(* IEC 61131-3 sources: JingjiangArm/moonboxpro_arm_8.4/Application/Application/任务列表/Main_Task, 12 files *)

(* ---- StErrParam_Use.st ---- *)
(*@CES
Name=StErrParam_Use
Type=Gvl
TypeGuid=2db5746d-d284-4425-9f7f-2663a34b0ebc
Guid=58394340-2af0-469d-907b-43e2b620f20c
HasDeclaration=True
HasImplementation=False
*)
{DECLARATION}
{attribute 'pack_mode' := '1'}
TYPE StErrParam_Use :(*这个是最终计算调整量需要的所有误差相关内容*)
STRUCT
	iErr_V: INT;(*纵向误差*)
	iErr_H: INT;(*横向误差*)
	iErr_V_Unprocessed	: INT;(*纵向误差-原始误差*)
	iErr_H_Unprocessed	: INT;(*横向误差-原始误差*)
	byIDX_V: BYTE;(*纵向索引*)
	byIDX_H: BYTE;(*横向索引*)
	byErrSts: BYTE;(*误差状态*)
	uiFSampleCounter:UINT;(*精采样数据计数*)
	iVerror_FollowPreUnit:INT;(*纵向跟踪前一色误差*)
	iVerror_Follow1Unit:INT;(*纵向跟踪第一色误差*)
	iHerror_FollowPreUnit :INT 	; (*横向跟前一色误差*)
	iHerror_Follow1Unit :INT 	;(*横向跟1色误差*)
	(*2025.9.16.094302*)
	iResult_VFollowpre_1stDerivate	: INT;(*YZJ计算误差*)
	//2025.11.13.105908||上传基线和峰值
	uiPeakValue_t1				: UINT;
	uiPeakValue_t2				: UINT;
	uiBaseUse_t1				: UINT;
	uiBaseUse_t2				: UINT;
	//2026.4.11.153149+2026.5.9.110438
	iErr_V_Display	: INT;(*纵向误差-显示平均处理*)
	iErr_H_Display	: INT;(*横向误差-原始误差*)

//2026.5.12.202228
	(*2026.5.10.150407/han.dp*)
	uiV_cam_raw: UINT;(*相机纵向原始误差*)
	iV_cam_pure: INT;(*相机纵向纯误差*)
	uiH_cam_raw: UINT;(*相机横向原始误差*)
	iH_cam_pure: INT;(*相机横向纯误差*)

END_STRUCT
END_TYPE

{IMPLEMENTATION}

(* ---- StTaskCycleDetection.st ---- *)
(*@CES
Name=StTaskCycleDetection
Type=Gvl
TypeGuid=2db5746d-d284-4425-9f7f-2663a34b0ebc
Guid=d17a89bb-f73c-4312-a6cf-f8b703e65793
HasDeclaration=True
HasImplementation=False
*)
{DECLARATION}
TYPE StTaskCycleDetection :
STRUCT
	xRstDetection			: BOOL;(* 复位测量 *)
	udiCycleCnt				: UDINT;(* 周期计数 *)
	xCalcIntervalEnabled	: BOOL;(* 计算间隔有效 *)
	tmTskIn					: TIME;(* 进入任务的时间戳 *)
	tmTskOut				: TIME;(* 离开任务的时间戳 *)
	tmTskIn_Prev			: TIME;(* 上次进入任务的时间戳 *)
	tmElapsed				: TIME;(* 任务消耗时间 *)
	tmElapsedMax			: TIME;(* 任务消耗时间最大 *)
	tmInterval				: TIME;(* 任务间隔 *)
	tmIntervalMax			: TIME;(* 任务间隔最大 *)
END_STRUCT
END_TYPE

{IMPLEMENTATION}

(* ---- KS_FlyMedian.st ---- *)
(*@CES
Name=KS_FlyMedian
Type=FunctionBlock
TypeGuid=6f9dac99-8de1-4efc-8465-68ac443b7d08
Guid=38054e60-5949-4eec-bd09-7b0f80079a4b
HasDeclaration=True
HasImplementation=True
*)
{DECLARATION}
FUNCTION KS_FlyMedian : REAL
(*中位数:与Python statistics.median语义一致——奇数取正中,偶数取中间两值的平均*)
(*插入排序会打乱入参缓冲区,窗口<=64,代价可忽略|Yang.zj+用于新飞点检测 2026.10.24.191149*)
VAR_INPUT
	pBuf	: POINTER TO REAL;(*缓冲区指针*)
	iCnt	: INT;			(*元素个数*)
END_VAR
VAR
	i		: INT;
	j		: INT;
	rTmp	: REAL;
END_VAR

{IMPLEMENTATION}
IF iCnt <= 0 THEN
	KS_FlyMedian:= 0.0;
	RETURN;
END_IF
FOR i:= 1 TO iCnt-1 DO(*插入排序*)
	rTmp:= pBuf[i];
	j:= i-1;
	WHILE (j >= 0) DO
		IF pBuf[j] > rTmp THEN
			pBuf[j+1]:= pBuf[j];
			j:= j-1;
		ELSE
			EXIT;
		END_IF
	END_WHILE
	pBuf[j+1]:= rTmp;
END_FOR
IF (iCnt MOD 2) = 1 THEN
	KS_FlyMedian:= pBuf[iCnt/2];
ELSE
	KS_FlyMedian:= (pBuf[iCnt/2-1] + pBuf[iCnt/2]) * 0.5;
END_IF

(* ---- KS_TskCycle_Begin.st ---- *)
(*@CES
Name=KS_TskCycle_Begin
Type=FunctionBlock
TypeGuid=6f9dac99-8de1-4efc-8465-68ac443b7d08
Guid=4df1a699-322b-4ad9-8d1d-9083be64c28d
HasDeclaration=True
HasImplementation=True
*)
{DECLARATION}
FUNCTION KS_TskCycle_Begin : INT
VAR_INPUT
	i_pstStTaskCycleDetection: POINTER TO StTaskCycleDetection;
END_VAR
VAR
	iResult: INT;
END_VAR
{IMPLEMENTATION}
iResult:= 0;
IF i_pstStTaskCycleDetection<>0 THEN
	i_pstStTaskCycleDetection^.tmTskIn:= TIME(); (* 进入的时间 *)
	i_pstStTaskCycleDetection^.udiCycleCnt:= i_pstStTaskCycleDetection^.udiCycleCnt+1; (* 进入一次就累计1次 *)
ELSE
	iResult:= -1;
END_IF
KS_TskCycle_Begin:= iResult;

(* ---- KS_TskCycle_End.st ---- *)
(*@CES
Name=KS_TskCycle_End
Type=FunctionBlock
TypeGuid=6f9dac99-8de1-4efc-8465-68ac443b7d08
Guid=379e6dd0-0b0c-44de-a9dc-120ed630a8f7
HasDeclaration=True
HasImplementation=True
*)
{DECLARATION}
FUNCTION KS_TskCycle_End : INT
VAR_INPUT
	i_pstStTaskCycleDetection: POINTER TO StTaskCycleDetection;
END_VAR
VAR
	iResult: INT;
END_VAR
{IMPLEMENTATION}
iResult:= 0;
IF i_pstStTaskCycleDetection<>0 THEN
	i_pstStTaskCycleDetection^.tmTskOut:= TIME(); (* 结束的时间 *)
	i_pstStTaskCycleDetection^.tmElapsed:= i_pstStTaskCycleDetection^.tmTskOut-i_pstStTaskCycleDetection^.tmTskIn; (* 算出本次耗时 *)
	IF i_pstStTaskCycleDetection^.tmElapsed>i_pstStTaskCycleDetection^.tmElapsedMax THEN (* 如果最高纪录有变化 *)
		i_pstStTaskCycleDetection^.tmElapsedMax:= i_pstStTaskCycleDetection^.tmElapsed;
	END_IF
	IF NOT i_pstStTaskCycleDetection^.xCalcIntervalEnabled THEN
		i_pstStTaskCycleDetection^.xCalcIntervalEnabled:= TRUE;
	ELSE
		i_pstStTaskCycleDetection^.tmInterval:= i_pstStTaskCycleDetection^.tmTskIn-i_pstStTaskCycleDetection^.tmTskIn_Prev; (* 周期间隔 *)
		IF i_pstStTaskCycleDetection^.tmInterval>i_pstStTaskCycleDetection^.tmIntervalMax THEN (* 如果周期间隔纪录有变化 *)
			i_pstStTaskCycleDetection^.tmIntervalMax:= i_pstStTaskCycleDetection^.tmInterval;
		END_IF
	END_IF

	i_pstStTaskCycleDetection^.tmTskIn_Prev:= i_pstStTaskCycleDetection^.tmTskIn; (* 上次进入的时间 *)

	IF i_pstStTaskCycleDetection^.xRstDetection THEN (* 重新计算周期的操作 *)
		i_pstStTaskCycleDetection^.xRstDetection:= FALSE;
		i_pstStTaskCycleDetection^.xCalcIntervalEnabled:= FALSE;
		i_pstStTaskCycleDetection^.tmElapsedMax:= T#0ms;
		i_pstStTaskCycleDetection^.tmIntervalMax:= T#0ms;
	END_IF
ELSE
	iResult:= -1;
END_IF

KS_TskCycle_End:= iResult;

(* ---- KS_UnPack_VisionERR.st ---- *)
(*@CES
Name=KS_UnPack_VisionERR
Type=FunctionBlock
TypeGuid=6f9dac99-8de1-4efc-8465-68ac443b7d08
Guid=46688986-88ab-493d-84a0-0feefd58abe3
HasDeclaration=True
HasImplementation=True
*)
{DECLARATION}
FUNCTION KS_UnPack_VisionERR : INT
VAR_INPUT
	i_wERR: WORD;(*接收到的误差值-加密数据*)
	i_pxFlag_valid: POINTER TO BOOL;(*bit15/有效标志*)
	i_pxFlag_update: POINTER TO BOOL;(*bit14/更新标志*)
	i_pxFlag_bitchk: POINTER TO BOOL;(*bit13/校验位*)
	i_piErr: POINTER TO INT;(*bit12~0/误差*)
END_VAR
VAR
	iRtn: INT := 0;(*默认0*)
END_VAR

{IMPLEMENTATION}
IF i_pxFlag_valid<>0 AND
	i_pxFlag_update<>0 AND
	i_pxFlag_bitchk<>0 AND
	i_piErr<>0 THEN
	iRtn:= 0;
	i_pxFlag_valid^:= WORD_TO_BOOL(SHR(i_wERR, 15) AND 16#1);
	i_pxFlag_update^:= WORD_TO_BOOL(SHR(i_wERR, 14) AND 16#1);
	i_pxFlag_bitchk^:= WORD_TO_BOOL(SHR(i_wERR, 13) AND 16#1);
	i_piErr^:= SHR(WORD_TO_INT(SHL(i_wERR, 3)), 3);
ELSE
	iRtn:= -1;
END_IF
KS_UnPack_VisionERR:= iRtn;

(* ---- KS_FB_AverageErr_Arc.st ---- *)
(*@CES
Name=KS_FB_AverageErr_Arc
Type=FunctionBlock
TypeGuid=6f9dac99-8de1-4efc-8465-68ac443b7d08
Guid=91f3b4d4-1a1f-49cc-9d09-db86b76ec74e
HasDeclaration=True
HasImplementation=True
*)
{DECLARATION}
FUNCTION_BLOCK KS_FB_AverageErr_Arc
VAR_INPUT
	i_xEn: BOOL;
	i_iErr: INT;(*输入的有效误差*)
	i_xErrValid: BOOL;(*误差有效性*)
	i_byAverageNum: BYTE;(*误差平均次数*)
END_VAR
VAR_OUTPUT
	o_xEn: BOOL;
	o_iErNo: INT;
	o_iErrResult: INT;
END_VAR
VAR
	rErrResult: REAL;(*误差平均使用的*)
	iBufferedIndexRd				: INT							;(*buffered array read index|*)
	iBufferedIndexWr				: INT							;(*buffered array write index|*)
	iPushedErrItemsAtLeast			: INT							;
	arErrorBuffered			: ARRAY [1..20] OF REAL						;
	iCountForSignalLost				: INT	;
	rSumTotal						: REAL;
	iIndex							: INT;
END_VAR

{IMPLEMENTATION}
o_xEn:= i_xEn;
o_iErNo:= 0;
IF i_xEn THEN
	IF i_byAverageNum>0 THEN
		rErrResult:= INT_TO_REAL(i_iErr);
		IF i_xErrValid THEN
			iBufferedIndexWr:= iBufferedIndexWr+1;
			IF iBufferedIndexWr>20 THEN
				iBufferedIndexWr:= iBufferedIndexWr-20;
			END_IF
			arErrorBuffered[iBufferedIndexWr]:= rErrResult;
			IF iPushedErrItemsAtLeast<i_byAverageNum THEN
				iPushedErrItemsAtLeast:= iPushedErrItemsAtLeast+1;
			ELSE
				IF i_byAverageNum>1 THEN
					iBufferedIndexRd:= iBufferedIndexWr;
					rSumTotal:= 0;
					FOR iIndex:=1 TO i_byAverageNum BY 1 DO
						rSumTotal:= rSumTotal+arErrorBuffered[iBufferedIndexRd];
						iBufferedIndexRd:= iBufferedIndexRd-1;
						IF iBufferedIndexRd<1 THEN
							iBufferedIndexRd:= iBufferedIndexRd+20;
						END_IF
					END_FOR
					rErrResult:= rSumTotal/i_byAverageNum;
				END_IF
			END_IF
			iCountForSignalLost:= 0;
			o_iErrResult:= REAL_TO_INT(rErrResult) ;
		ELSE(*连续丢失3幅就重新开始计算平均*)
			iCountForSignalLost:= 	iCountForSignalLost+1;
			IF 	iCountForSignalLost>3 THEN
				iBufferedIndexWr:= 0;
				iPushedErrItemsAtLeast:= 0;
			END_IF
			o_iErNo:= -1;
		END_IF
	ELSE
		o_iErrResult:= i_iErr;
	END_IF
END_IF

(* ---- KS_FB_GetError_Arc.st ---- *)
(*@CES
Name=KS_FB_GetError_Arc
Type=FunctionBlock
TypeGuid=6f9dac99-8de1-4efc-8465-68ac443b7d08
Guid=34f07fc4-d98c-4616-a827-05a7c8017d66
HasDeclaration=True
HasImplementation=True
*)
{DECLARATION}
FUNCTION_BLOCK KS_FB_GetError_Arc
VAR_INPUT
	i_xEn: BOOL;
	i_iUnitMax: INT;
	i_byGetErrMode: BYTE;(*获取误差方式，
	1：读取金刚来的误差
	2：读取月光宝盒/月光宝盒PRO来的误差
	*)
	i_aiAlarm_V: ARRAY [1..MAX_UNIT_NUM] OF INT;(*后续换成全局输入的变量*)
	i_aiAlarm_H: ARRAY [1..MAX_UNIT_NUM] OF INT;(*后续换成全局输入的变量*)
	i_aiAdjust_V: ARRAY [1..MAX_UNIT_NUM] OF INT;(*修正量*)
	i_aiAdjust_H: ARRAY [1..MAX_UNIT_NUM] OF INT;(*修正量*)

	i_abyAverageNum_V: ARRAY [1..MAX_UNIT_NUM] OF BYTE;(*误差平均次数*)
	i_abyAverageNum_H: ARRAY [1..MAX_UNIT_NUM] OF BYTE;(*误差平均次数*)
	//2026.4.11.150236 误差显示平均
	i_abyAverageNum_V_Display: ARRAY [1..MAX_UNIT_NUM] OF BYTE;(*误差显示平均次数*)
	i_abyAverageNum_H_Display: ARRAY [1..MAX_UNIT_NUM] OF BYTE;(*误差显示平均次数*)
	i_pstStSysParam								: POINTER TO StSysParam;
END_VAR
VAR_OUTPUT
	o_xEn: BOOL;
	o_iNoEr: INT;
	o_astStErrParam_Use: ARRAY [1..MAX_UNIT_NUM] OF StErrParam_Use;
END_VAR
VAR
	iN: INT;
	aiError_and_Sts_V: ARRAY [1..MAX_UNIT_NUM] OF INT;(*读取的来自金刚/月光宝盒PRO的误差及状态*)
	aiError_and_Sts_H: ARRAY [1..MAX_UNIT_NUM] OF INT;(*读取的来自金刚/月光宝盒PRO的误差及状态*)
	iTemp: WORD;
	aiError_V: ARRAY [1..MAX_UNIT_NUM] OF INT;(*处理完成后的纵向误差列表*)
	aiError_H: ARRAY [1..MAX_UNIT_NUM] OF INT;(*处理完成后的横向误差列表*)
	abyErrSts: ARRAY [1..MAX_UNIT_NUM] OF BYTE;(*处理完成后的纵横向误差状态*)
	abyIndex_V: ARRAY [1..MAX_UNIT_NUM] OF BYTE;(*处理完成后的索引*)
	abyIndex_H: ARRAY [1..MAX_UNIT_NUM] OF BYTE;(*处理完成后的索引*)
	axValid_V: ARRAY [1..MAX_UNIT_NUM] OF BOOL;(*误差有效性*)
	axValid_H: ARRAY [1..MAX_UNIT_NUM] OF BOOL;(*误差有效性*)
	axFlag_Refresh_V: ARRAY [1..MAX_UNIT_NUM] OF BOOL;(*误差刷新标志*)
	axFlag_Refresh_H: ARRAY [1..MAX_UNIT_NUM] OF BOOL;(*误差刷新标志*)
	axFlag_Check_V: ARRAY [1..MAX_UNIT_NUM] OF BOOL;(*误差校验位*)
	axFlag_Check_H: ARRAY [1..MAX_UNIT_NUM] OF BOOL;(*误差校验位*)
	axFlag_PreRefresh_V: ARRAY [1..MAX_UNIT_NUM] OF BOOL;(*误差有效性*)
	axFlag_PreRefresh_H: ARRAY [1..MAX_UNIT_NUM] OF BOOL;(*误差有效性*)
	afbKS_FB_PickOutFakePoint_V: ARRAY [1..MAX_UNIT_NUM] OF KS_FB_PickOutFakePoint;(*误差飞点处理*)
	afbKS_FB_PickOutFakePoint_H: ARRAY [1..MAX_UNIT_NUM] OF KS_FB_PickOutFakePoint;
	afbKS_FB_AverageErr_Arc_V: ARRAY [1..MAX_UNIT_NUM] OF KS_FB_AverageErr_Arc;(*误差平均处理*)
	afbKS_FB_AverageErr_Arc_H: ARRAY [1..MAX_UNIT_NUM] OF KS_FB_AverageErr_Arc;
	//2026.4.11.150050+
	afbKS_FB_AverageErr_Arc_V_Display: ARRAY [1..MAX_UNIT_NUM] OF KS_FB_AverageErr_Arc;(*误差平均处理@界面显示*)
	afbKS_FB_AverageErr_Arc_H_Display: ARRAY [1..MAX_UNIT_NUM] OF KS_FB_AverageErr_Arc;

	aiError_V_Res_Display: ARRAY [1..MAX_UNIT_NUM] OF INT;(*处理完成后的纵向显示误差列表*)
	aiError_H_Res_Display: ARRAY [1..MAX_UNIT_NUM] OF INT;(*处理完成后的横向显示误差列表*)
	//2026.5.9.110955
	axFakePoint_V: ARRAY [1..MAX_UNIT_NUM] OF BOOL;
	axFakePoint_H: ARRAY [1..MAX_UNIT_NUM] OF BOOL;

	aiError_V_Res: ARRAY [1..MAX_UNIT_NUM] OF INT;(*处理完成后的纵向误差列表*)
	aiError_H_Res: ARRAY [1..MAX_UNIT_NUM] OF INT;(*处理完成后的横向误差列表*)
	abyIndex_V_Pre: ARRAY [1..MAX_UNIT_NUM] OF BYTE;(*处理完成后的索引*)
	abyIndex_H_Pre: ARRAY [1..MAX_UNIT_NUM] OF BYTE;(*处理完成后的索引*)
	iUnitNR: INT;
	iStationId: INT;
	dwOFST2: DWORD;
	iRtn: INT;
	stStProtocol_PDU_Up_Rd: StParam_PDU_Up;
	pstStCMD_F05_: POINTER TO StPdu_Up_05;
	pbyTemp: POINTER TO BYTE;
	wCHK_Up_Calc: WORD;
	dwCheckSumVal: DWORD;
	abyBuf_PduCmd_rcv: ARRAY [1..MAX_PDU_CMD_BYTES_UP] OF BYTE; (* 2021.12.4.163129/hdp/读取 *)
	xtest: BOOL;
	aiResult_VFollowpre_1stDerivate: ARRAY [1..MAX_UNIT_NUM] OF INT;

	//alTime: ARRAY [1..10] OF LTIME;
	abyBuf_PduCmd_rcv_All: ARRAY [1..1000] OF BYTE;

	//新飞点剔除:每色组纵横各一个独立实例(总开关gc_xUseNewFlyRemove在GCL)|Yang.zj+用于新飞点检测 2026.10.24.191149
	afbKS_FlyRemove_V: ARRAY [1..MAX_UNIT_NUM] OF KS_FlyRemove;
	afbKS_FlyRemove_H: ARRAY [1..MAX_UNIT_NUM] OF KS_FlyRemove;
	aiError_V_Fly: ARRAY [1..MAX_UNIT_NUM] OF INT;(*剔除后送平均的纵向误差*)
	aiError_H_Fly: ARRAY [1..MAX_UNIT_NUM] OF INT;(*剔除后送平均的横向误差*)
	xFlyNewFrame: BOOL;(*本周期该色组是否来了新帧*)
	xFlyReset: BOOL;(*该色组剔除器复位请求*)
	aiFlyMarkModePre: ARRAY [1..MAX_UNIT_NUM] OF INT;(*上次色标排列模式*)
	abyFlySignalPre: ARRAY [1..MAX_UNIT_NUM] OF BYTE;(*上次RGB信号通道*)
	axFlyHorEnPre: ARRAY [1..MAX_UNIT_NUM] OF BOOL;(*上次横向开关*)
END_VAR

{IMPLEMENTATION}
o_xEn:= i_xEn;
o_iNoEr:= 0;
IF i_xEn THEN
	IF i_iUnitMax>0 THEN
	CASE i_byGetErrMode OF
			1:
				FOR iN:=1 TO i_iUnitMax BY 1 DO
					iTemp:= aiError_and_Sts_V[iN];
					axValid_V[iN]:= INT_TO_BOOL(iTemp AND 16#04);(*bit2:有效位*)
					axFlag_Refresh_V[iN]:= INT_TO_BOOL(iTemp AND 16#02);(*bit1:刷新位*)
					axFlag_Check_V[iN]:= INT_TO_BOOL(iTemp AND 16#01);(*bit0:校验位*)
					IF axFlag_PreRefresh_V[iN]<>axFlag_Refresh_V[iN] THEN	 	(*误差已刷新*)
						IF axValid_V[iN] THEN
							aiError_V[iN]:= SHR(iTemp,3);(*误差*)
						ELSE
							aiError_V[iN]:= gc_iValueReferToLost;
							abyErrSts[iN].1:= TRUE;(*纵向丢失*)
						END_IF
						abyIndex_V[iN]:= abyIndex_V[iN]+1;
					END_IF
					axFlag_PreRefresh_V[iN]:= axFlag_Refresh_V[iN];
					(*纵向误差处理完成*)
					iTemp:= aiError_and_Sts_H[iN];
					axValid_H[iN]:= INT_TO_BOOL(iTemp AND 16#04);(*bit2:有效位*)
					axFlag_Refresh_H[iN]:= INT_TO_BOOL(iTemp AND 16#02);(*bit1:刷新位*)
					axFlag_Check_H[iN]:= INT_TO_BOOL(iTemp AND 16#01);(*bit0:校验位*)
					IF axFlag_PreRefresh_H[iN]<>axFlag_Refresh_H[iN] THEN	 	(*误差已刷新*)
						IF axValid_H[iN] THEN
							aiError_H[iN]:= SHR(iTemp,3);(*误差*)
						ELSE
							aiError_H[iN]:= gc_iValueReferToLost;
							abyErrSts[iN].5:= TRUE;(*横向丢失*)
						END_IF
						abyIndex_H[iN]:= abyIndex_H[iN]+1;
					END_IF
					axFlag_PreRefresh_H[iN]:= axFlag_Refresh_H[iN];
					(*横向误差处理完成*)
				END_FOR
			2:
				//alTime[4] := LTIME();
				dwOFST2:= 0;
				iRtn := GTN_RN_UserPCRdLocalFPGA(
							1,1,
							0,//0,
							ADR(abyBuf_PduCmd_rcv_All),
							DWORD_TO_WORD(dwOFST2),
							KS_GetNumOfDwordUsed(INT_TO_DWORD(i_iUnitMax)*MAX_PDU_CMD_BYTES_DN));
				FOR iN:=1 TO i_iUnitMax BY 1 DO
					iUnitNR:= iN;(*通讯轴号也需要根据后续系统配置处理*)
					iStationId:= g_stStSysParam.stStSysParam_UnSave.aiStationList_UnitController[iN];(*2024.1.3.200541/+ *)
					IF KS_IsValidStationNR(iStationId) THEN
					(*读取从站即时上报的数据|每次32Bytes|*)
//2025.11.20.172237
//						dwOFST2 := MAX_PDU_CMD_BYTES_DN*(iUnitNR-1);
// 						dwOFST2.14:= TRUE;(* 绝对地址访问 *)
(*						iRtn := GTN_RN_UserPCRdLocalFPGA(1,1,
									0,//INT_TO_BYTE(iStationId),
									ADR(stStProtocol_PDU_Up_Rd),
									DWORD_TO_WORD(dwOFST2),
									15);//16448
									*)
// 						iRtn := GTN_RN_UserPCRdLocalFPGA(
// 									ADR(stStProtocol_PDU_Up_Rd),
// 									0,//INT_TO_BYTE(iStationId),
// 									DWORD_TO_WORD(dwOFST2),
// 									15);//16448

//2025.11.20.172246
//						iRtn := GTN_RN_UserPCRdLocalFPGA(
// 									1,1,
// 									0,//0,
// 									ADR(abyBuf_PduCmd_rcv),
// 									DWORD_TO_WORD(dwOFST2),
// 									15);//16448
					dwOFST2 := MAX_PDU_CMD_BYTES_DN*(iUnitNR-1);

					SysMemCpy(ADR(stStProtocol_PDU_Up_Rd),ADR(abyBuf_PduCmd_rcv_All)+dwOFST2,SIZEOF(stStProtocol_PDU_Up_Rd));
					(*检查命令|*)
						pstStCMD_F05_:=0;

						pbyTemp:= ADR(stStProtocol_PDU_Up_Rd.byPkgId);
						wCHK_Up_Calc:= KS_CRC(pbyTemp, 46, ADR(dwCheckSumVal));(*51是wCHK之前的数据长度*)
						IF wCHK_Up_Calc=stStProtocol_PDU_Up_Rd.wCHK THEN (*CRC校验通过*)
							CASE stStProtocol_PDU_Up_Rd.byPkgId OF
								5:
								pstStCMD_F05_:= ADR(stStProtocol_PDU_Up_Rd.abyPayload);
								IF pstStCMD_F05_<>0 THEN
									aiError_V[iN]:= stStProtocol_PDU_Up_Rd.iErr_V_Raw;
									aiError_H[iN]:= stStProtocol_PDU_Up_Rd.iErr_H_Raw;
									abyIndex_V[iN]:= stStProtocol_PDU_Up_Rd.byIDX_V;
									abyIndex_H[iN]:= stStProtocol_PDU_Up_Rd.byIDX_H;
									IF aiError_V[iN]=gc_iValueReferToLost THEN
										abyErrSts[iN].1:= TRUE;(*纵向丢失*)
									ELSE
										axValid_V[iN]:= TRUE;
									END_IF
									IF aiError_H[iN]=gc_iValueReferToLost THEN
										abyErrSts[iN].5:= TRUE;(*横向丢失*)
									ELSE
										axValid_H[iN]:= TRUE;
									END_IF
									o_astStErrParam_Use[iN].iResult_VFollowpre_1stDerivate:=
											pstStCMD_F05_^.iResult_VFollowpre_1stDerivate;
									aiResult_VFollowpre_1stDerivate[iN]:=
											pstStCMD_F05_^.iResult_VFollowpre_1stDerivate;
									//2025.11.13.110235上传基线和峰值
									o_astStErrParam_Use[iN].uiBaseUse_t1:= pstStCMD_F05_^.uiBaseUse_t1;
									o_astStErrParam_Use[iN].uiBaseUse_t2:= pstStCMD_F05_^.uiBaseUse_t2;
									o_astStErrParam_Use[iN].uiPeakValue_t1:= pstStCMD_F05_^.uiPeakValue_t1;
									o_astStErrParam_Use[iN].uiPeakValue_t2:= pstStCMD_F05_^.uiPeakValue_t2;
								//2026.5.9.110642
									i_pstStSysParam^.astStRSV_UnitParam_UnSave[iN].iCurLabelPos:= pstStCMD_F05_^.iCurLabelPos;(*本色三角标位置，点数*)
									i_pstStSysParam^.astStRSV_UnitParam_UnSave[iN].iPreLabelPos:= pstStCMD_F05_^.iPreLabelPos;(*前色三角标位置，点数*)
									i_pstStSysParam^.astStRSV_UnitParam_UnSave[iN].byFlag_CommFromSlave:= pstStCMD_F05_^.byFlag_CommFromSlave;(*bit0 xFlag_FindFirstSuccess;bit1 xFlag_FindPreSuccess*)
									i_pstStSysParam^.astStRSV_UnitParam_UnSave[iN].xFlag_FindFirstSuccess:= i_pstStSysParam^.astStRSV_UnitParam_UnSave[iN].byFlag_CommFromSlave.0;
									i_pstStSysParam^.astStRSV_UnitParam_UnSave[iN].xFlag_FindPreSuccess:= i_pstStSysParam^.astStRSV_UnitParam_UnSave[iN].byFlag_CommFromSlave.1;
									i_pstStSysParam^.astStRSV_UnitParam_UnSave[iN].byDetectedSignalCount:= pstStCMD_F05_^.byDetectedSignalCount;(*当前检测到色标个数*)
									i_pstStSysParam^.astStRSV_UnitParam_UnSave[iN].byMarkStep:= pstStCMD_F05_^.byMarkStep;(*当前全自动套印步骤*)
									i_pstStSysParam^.astStRSV_UnitParam_UnSave[iN].rGateSignalWidth_R:= BYTE_TO_REAL (pstStCMD_F05_^.byWidthRS) /10.0;(*粗采样计算波形宽度*)

								END_IF
							END_CASE
						END_IF
					END_IF
				END_FOR

			ELSE
			(*其他状态时，就先按丢失处理*)
				FOR iN:=1 TO MAX_UNIT_NUM BY 1 DO
					aiError_V[iN]:= gc_iValueReferToLost;
					aiError_H[iN]:= gc_iValueReferToLost;
					abyErrSts[iN].1:= TRUE;(*纵向丢失*)
					abyErrSts[iN].5:= TRUE;(*横向丢失*)
				END_FOR
		END_CASE

		(*从这里开始进行误差处理-飞点和平均*)
		(*飞点处理*)

		(*FOR iN:=1 TO MAX_UNIT_NUM BY 1 DO
			IF abyIndex_V_Pre[iN]<>abyIndex_V[iN] AND abyIndex_H_Pre[iN]<>abyIndex_H[iN] THEN
				abyErrSts[iN]:= 0;
				axValid_V[iN]:= FALSE;
				axValid_H[iN]:= FALSE;
				IF aiError_V[iN]=gc_iValueReferToLost THEN
					abyErrSts[iN].1:= TRUE;(*纵向丢失*)
				ELSE
					axValid_V[iN]:= TRUE;
				END_IF
				IF aiError_H[iN]=gc_iValueReferToLost THEN
					abyErrSts[iN].5:= TRUE;(*横向丢失*)
				ELSE
					axValid_H[iN]:= TRUE;
				END_IF
				o_astStErrParam_Use[iN].iResult_VFollowpre_1stDerivate:=
						aiResult_VFollowpre_1stDerivate[iN];

				o_astStErrParam_Use[iN].byIDX_V:= abyIndex_V[iN];
				o_astStErrParam_Use[iN].byIDX_H:= abyIndex_H[iN];
	//2026.02.08.195855
				(*平均处理*)
				afbKS_FB_AverageErr_Arc_V[iN](
					i_xEn:= TRUE,
					i_iErr:= aiError_V[iN],
					i_xErrValid:= axValid_V[iN],(*2025.01.03.110017*)
					i_byAverageNum:= i_abyAverageNum_V[iN],
					o_iErrResult=>aiError_V_Res[iN]);
				axFakePoint_V[iN]:= FALSE;

				afbKS_FB_PickOutFakePoint_V[iN](
					i_xIsValidError:= axValid_V[iN],
					i_iError_0_01mm:= aiError_V_Res[iN],
					i_iVariationBaseValue:= 50,(*2025.01.03.110017*)
					i_iBoundaryError_0_01mm:= 20,
					i_iErrorLevel_0_01mm:= 25,
					i_iVariationVariationMin:= 5,
					i_iVariationVariationMax:= 50,
					o_xFakeIsConfirmed=> axFakePoint_V[iN]);
	//2026.02.08.195945
				afbKS_FB_AverageErr_Arc_H[iN](
					i_xEn:= TRUE,
					i_iErr:= aiError_H[iN],
					i_xErrValid:= axValid_H[iN],(*2025.01.03.110017*)
					i_byAverageNum:= i_abyAverageNum_H[iN],
					o_iErrResult=>aiError_H_Res[iN]);
				axFakePoint_H[iN]:= FALSE;

				afbKS_FB_PickOutFakePoint_H[iN](
					i_xIsValidError:= axValid_H[iN],
					i_iError_0_01mm:= aiError_H_Res[iN],
					i_iVariationBaseValue:= 50,
					i_iBoundaryError_0_01mm:= 20,
					i_iErrorLevel_0_01mm:= 25,
					i_iVariationVariationMin:= 5,
					i_iVariationVariationMax:= 50,
					o_xFakeIsConfirmed=> axFakePoint_H[iN]);

				//显示平均@2026.4.11.150119+
				afbKS_FB_AverageErr_Arc_V_Display[iN](
					i_xEn:= TRUE,
					i_iErr:= aiError_V[iN],
					i_xErrValid:= axValid_V[iN],(*2025.01.03.110017*)
					i_byAverageNum:= i_abyAverageNum_V_Display[iN],
					o_iErrResult=>aiError_V_Res_Display[iN]);

				afbKS_FB_AverageErr_Arc_H_Display[iN](
					i_xEn:= TRUE,
					i_iErr:= aiError_H[iN],
					i_xErrValid:= axValid_H[iN],(*2025.01.03.110017*)
					i_byAverageNum:= i_abyAverageNum_H_Display[iN],
					o_iErrResult=>aiError_H_Res_Display[iN]);

			END_IF*)
		FOR iN:=1 TO MAX_UNIT_NUM BY 1 DO
			(*新飞点剔除:误差平均之前对原始逐帧误差剔除,成熟账本时为外推 P 并刷锁存，否则锁存,必须先剔除再平均,否则飞点被N幅平均稀释后可能低于门限漏掉*)
			(*总开关gc_xUseNewFlyRemove在GCL,置FALSE并重编译即回退旧逻辑;飞点/暂缓帧置axFakePoint_V/H(byErrSts.2/6),阶跃(真实变化)不置位|Yang.zj+用于新飞点检测 2026.10.24.191149*)
			IF gc_xUseNewFlyRemove THEN
				xFlyNewFrame:= (abyIndex_V_Pre[iN]<>abyIndex_V[iN]) AND (abyIndex_H_Pre[iN]<>abyIndex_H[iN]);
				(*工况切换检测:色标排列模式/RGB信号通道/横向开关任一变化,该色组剔除器可信历史不可信,复位重新暖机*)
				xFlyReset:= FALSE;
				IF i_pstStSysParam<>0 THEN
					IF (aiFlyMarkModePre[iN]<>i_pstStSysParam^.astStUnitParam_Save[iN].iMarkArrangeMode)
						OR (abyFlySignalPre[iN]<>i_pstStSysParam^.astStUnitParam_Save[iN].bySignalSelect)
						OR (axFlyHorEnPre[iN]<>i_pstStSysParam^.astStUnitParam_Save[iN].dwFlag_Ctl.0) THEN
						aiFlyMarkModePre[iN]:= i_pstStSysParam^.astStUnitParam_Save[iN].iMarkArrangeMode;
						abyFlySignalPre[iN]:= i_pstStSysParam^.astStUnitParam_Save[iN].bySignalSelect;
						axFlyHorEnPre[iN]:= i_pstStSysParam^.astStUnitParam_Save[iN].dwFlag_Ctl.0;
						xFlyReset:= TRUE;
					END_IF
				END_IF
				afbKS_FlyRemove_V[iN](
					i_iErr:= aiError_V[iN],
					i_xErrValid:= xFlyNewFrame AND (aiError_V[iN]<>gc_iValueReferToLost),
					i_xLost:= xFlyNewFrame AND (aiError_V[iN]=gc_iValueReferToLost),
					i_xReset:= xFlyReset,
					o_iErrResult=> aiError_V_Fly[iN],
					o_xFake=> axFakePoint_V[iN]);
				afbKS_FlyRemove_H[iN](
					i_iErr:= aiError_H[iN],
					i_xErrValid:= xFlyNewFrame AND (aiError_H[iN]<>gc_iValueReferToLost),
					i_xLost:= xFlyNewFrame AND (aiError_H[iN]=gc_iValueReferToLost),
					i_xReset:= xFlyReset,
					o_iErrResult=> aiError_H_Fly[iN],
					o_xFake=> axFakePoint_H[iN]);
			ELSE
				aiError_V_Fly[iN]:= aiError_V[iN];(*旧路径:不剔除,原值送平均*)
				aiError_H_Fly[iN]:= aiError_H[iN];
			END_IF
			IF abyIndex_V_Pre[iN]<>abyIndex_V[iN] AND abyIndex_H_Pre[iN]<>abyIndex_H[iN] THEN
				abyErrSts[iN]:= 0;
				axValid_V[iN]:= FALSE;
				axValid_H[iN]:= FALSE;
				IF aiError_V[iN]=gc_iValueReferToLost THEN
					abyErrSts[iN].1:= TRUE;(*纵向丢失*)
				ELSE
					axValid_V[iN]:= TRUE;
				END_IF
				IF aiError_H[iN]=gc_iValueReferToLost THEN
					abyErrSts[iN].5:= TRUE;(*横向丢失*)
				ELSE
					axValid_H[iN]:= TRUE;
				END_IF
				o_astStErrParam_Use[iN].iResult_VFollowpre_1stDerivate:=
						aiResult_VFollowpre_1stDerivate[iN];

				o_astStErrParam_Use[iN].byIDX_V:= abyIndex_V[iN];
				o_astStErrParam_Use[iN].byIDX_H:= abyIndex_H[iN];
//2026.02.08.195855
				(*平均处理*)
				afbKS_FB_AverageErr_Arc_V[iN](
					i_xEn:= TRUE,
					i_iErr:= aiError_V_Fly[iN],(*新飞点:喂剔除后的值|Yang.zj+用于新飞点检测 2026.10.24.191149*)
					i_xErrValid:= axValid_V[iN],(*2025.01.03.110017*)
					i_byAverageNum:= i_abyAverageNum_V[iN],
					o_iErrResult=>aiError_V_Res[iN]);
				IF NOT gc_xUseNewFlyRemove THEN(*旧飞点判断:新算法启用时整块跳过|Yang.zj+用于新飞点检测 2026.10.24.191149*)
				axFakePoint_V[iN]:= FALSE;

				afbKS_FB_PickOutFakePoint_V[iN](
					i_xIsValidError:= axValid_V[iN],
					i_iError_0_01mm:= aiError_V_Res[iN],
					i_iVariationBaseValue:= 50,(*2025.01.03.110017*)
					i_iBoundaryError_0_01mm:= 20,
					i_iErrorLevel_0_01mm:= 25,
					i_iVariationVariationMin:= 5,
					i_iVariationVariationMax:= 50,
					o_xFakeIsConfirmed=> axFakePoint_V[iN]);
				END_IF
//2026.02.08.195945
				afbKS_FB_AverageErr_Arc_H[iN](
					i_xEn:= TRUE,
					i_iErr:= aiError_H_Fly[iN],(*新飞点:喂剔除后的值|Yang.zj+用于新飞点检测 2026.10.24.191149*)
					i_xErrValid:= axValid_H[iN],(*2025.01.03.110017*)
					i_byAverageNum:= i_abyAverageNum_H[iN],
					o_iErrResult=>aiError_H_Res[iN]);
				IF NOT gc_xUseNewFlyRemove THEN(*旧飞点判断:新算法启用时整块跳过|Yang.zj+用于新飞点检测 2026.10.24.191149*)
				axFakePoint_H[iN]:= FALSE;

				afbKS_FB_PickOutFakePoint_H[iN](
					i_xIsValidError:= axValid_H[iN],
					i_iError_0_01mm:= aiError_H_Res[iN],
					i_iVariationBaseValue:= 50,
					i_iBoundaryError_0_01mm:= 20,
					i_iErrorLevel_0_01mm:= 25,
					i_iVariationVariationMin:= 5,
					i_iVariationVariationMax:= 50,
					o_xFakeIsConfirmed=> axFakePoint_H[iN]);
				END_IF

				//显示平均@2026.4.11.150119+
				afbKS_FB_AverageErr_Arc_V_Display[iN](
					i_xEn:= TRUE,
					i_iErr:= aiError_V_Fly[iN],(*新飞点:喂剔除后的值|Yang.zj+用于新飞点检测 2026.10.24.191149*)
					i_xErrValid:= axValid_V[iN],(*2025.01.03.110017*)
					i_byAverageNum:= i_abyAverageNum_V_Display[iN],
					o_iErrResult=>aiError_V_Res_Display[iN]);

				afbKS_FB_AverageErr_Arc_H_Display[iN](
					i_xEn:= TRUE,
					i_iErr:= aiError_H_Fly[iN],(*新飞点:喂剔除后的值|Yang.zj+用于新飞点检测 2026.10.24.191149*)
					i_xErrValid:= axValid_H[iN],(*2025.01.03.110017*)
					i_byAverageNum:= i_abyAverageNum_H_Display[iN],
					o_iErrResult=>aiError_H_Res_Display[iN]);
			END_IF
			(*到这里误差的飞点和平均都处理完了，该处理其他东西了*)
			o_astStErrParam_Use[iN].iErr_V_Unprocessed:= aiError_V[iN];(*原始误差*)
			o_astStErrParam_Use[iN].iErr_H_Unprocessed:= aiError_H[iN];
			o_astStErrParam_Use[iN].byErrSts:= 0;
			o_astStErrParam_Use[iN].byErrSts:= abyErrSts[iN];(*现在的状态*)

//2026.5.9.110835处理一下显示平均相关
			IF NOT o_astStErrParam_Use[iN].byErrSts.1 THEN(*纵向未丢失*)
				o_astStErrParam_Use[iN].iErr_V:= aiError_V_Res[iN]-i_aiAdjust_V[iN];
				//2026.4.11.150603+
				o_astStErrParam_Use[iN].iErr_V_Display:= aiError_V_Res_Display[iN]-i_aiAdjust_V[iN];
				IF axFakePoint_V[iN] THEN(*飞点*)
					o_astStErrParam_Use[iN].byErrSts.2:= TRUE;
				END_IF
				(*报警标志检查*)
				//IF ABS(o_astStErrParam_Use[iN].iErr_V)>ABS(i_aiAlarm_V[iN]) THEN
				IF ABS(o_astStErrParam_Use[iN].iErr_V_Display)>ABS(i_aiAlarm_V[iN]) THEN
					o_astStErrParam_Use[iN].byErrSts.0:= TRUE;
				END_IF
			ELSE
				o_astStErrParam_Use[iN].iErr_V:= gc_iValueReferToLost;
				o_astStErrParam_Use[iN].iErr_V_Display:= gc_iValueReferToLost;
			END_IF
			IF NOT o_astStErrParam_Use[iN].byErrSts.5 THEN(*横向未丢失*)
				o_astStErrParam_Use[iN].iErr_H:= aiError_H_Res[iN]-i_aiAdjust_H[iN];(*处理完的误差-修正量*)
				//2026.4.11.150603+
				o_astStErrParam_Use[iN].iErr_H_Display:= aiError_H_Res_Display[iN]-i_aiAdjust_H[iN];
				IF axFakePoint_H[iN] THEN(*飞点*)
					o_astStErrParam_Use[iN].byErrSts.6:= TRUE;
				END_IF
				(*报警标志检查*)
				//IF ABS(o_astStErrParam_Use[iN].iErr_H)>ABS(i_aiAlarm_H[iN]) THEN
				IF ABS(o_astStErrParam_Use[iN].iErr_H_Display)>ABS(i_aiAlarm_H[iN]) THEN
					o_astStErrParam_Use[iN].byErrSts.4:= TRUE;
				END_IF
			ELSE
				o_astStErrParam_Use[iN].iErr_H:= gc_iValueReferToLost;
				//2026.4.11.150603+
				o_astStErrParam_Use[iN].iErr_H_Display:= gc_iValueReferToLost;
			END_IF
			abyIndex_V_Pre[iN]:= abyIndex_V[iN];
			abyIndex_H_Pre[iN]:= abyIndex_H[iN];
		END_FOR
	END_IF
END_IF

(* ---- KS_FB_GetError_Arc_1.st ---- *)
(*@CES
Name=KS_FB_GetError_Arc_1
Type=FunctionBlock
TypeGuid=6f9dac99-8de1-4efc-8465-68ac443b7d08
Guid=a8fc5d1b-180f-4776-912e-45955a246124
HasDeclaration=True
HasImplementation=True
*)
{DECLARATION}
FUNCTION_BLOCK KS_FB_GetError_Arc_1
VAR_INPUT
	i_xEn: BOOL;(*该功能的使能条件*)
	i_iUnitMax: INT;(*有效色组范围1..MAX_UNIT_NUM*)
	i_abyGetErrMode: ARRAY [1..MAX_UNIT_NUM] OF BYTE;
	(*2026.5.10.102830/han.dp/修正接口定义方式:
	bit0 月光宝盒PRO误差源,1有效
	bit1 金刚误差源,1有效
	bit4 相机安装方向-反向/2026.5.24.173347/han.dp
	bit5 逆序/2026.5.24.173354/han.dp
	bit7 用于标记有效位标志; =0表示bit0有效,以月光宝盒PRO的误差作为调整依据; =1表示bit1有效,以金刚误差作为调整参考;
	--------------------------------------------------
	举例:
	* 16#01来自月光宝盒PRO;
	* 16#82来自视觉,并作为调整依据;
	* 16#03金刚和月光宝盒PRO误差都读,但只以月光宝盒PRO的误差作为调整依据;
	* 16#83金刚和月光宝盒PRO误差都读,但只以金刚的误差作为调整依据;
	*)
	i_aiAlarm_V: ARRAY [1..MAX_UNIT_NUM] OF INT;(*后续换成全局输入的变量*)
	i_aiAlarm_H: ARRAY [1..MAX_UNIT_NUM] OF INT;(*后续换成全局输入的变量*)
	i_aiAdjust_V: ARRAY [1..MAX_UNIT_NUM] OF INT;(*修正量*)
	i_aiAdjust_H: ARRAY [1..MAX_UNIT_NUM] OF INT;(*修正量*)
	i_abyAverageNum_V: ARRAY [1..MAX_UNIT_NUM] OF BYTE;(*误差平均次数*)
	i_abyAverageNum_H: ARRAY [1..MAX_UNIT_NUM] OF BYTE;(*误差平均次数*)
	(*统一注释0916+2026.4.11.150236 误差显示平均*)
	i_abyAverageNum_V_Display: ARRAY [1..MAX_UNIT_NUM] OF BYTE;(*误差显示平均次数*)
	i_abyAverageNum_H_Display: ARRAY [1..MAX_UNIT_NUM] OF BYTE;(*误差显示平均次数*)
	i_pstStSysParam								: POINTER TO StSysParam;
	i_dwKSMatrixMark: DWORD;(*2026.5.24.173538/han.dp/科赛矩阵色标描述/高16bit和低16bit分别为ab值*)
END_VAR
VAR_OUTPUT
	o_xEno: BOOL;
	o_iErNo: INT;
	o_astStErrParam_Use: ARRAY [1..MAX_UNIT_NUM] OF StErrParam_Use;
	o_stSystimeElapsed: SYSTIME;(*2026.5.24.152004/han.dp*)
END_VAR
VAR
	xInitialized_Ref_KSMatrixMark: BOOL := FALSE;
	abyGetErrMode_Ref: ARRAY [1..MAX_UNIT_NUM] OF BYTE := [0];
	dwKSMatrixMark_Ref: DWORD := 0;
	aiRef_KSMatrixMark: ARRAY [1..MAX_UNIT_NUM,1..2] OF INT;(*16色色标的参考位置*)
	wKSMatrixMark_Hword: WORD;
	wKSMatrixMark_Lword: WORD;

	iN: INT;
	aiError_and_Sts_V: ARRAY [1..MAX_UNIT_NUM] OF INT;(*读取的来自金刚/月光宝盒PRO的误差及状态*)
	aiError_and_Sts_H: ARRAY [1..MAX_UNIT_NUM] OF INT;(*读取的来自金刚/月光宝盒PRO的误差及状态*)
	iTemp: WORD;

(*deprecated@2026.5.28.172423/han.dp
	axFlag_Refresh_V: ARRAY [1..MAX_UNIT_NUM] OF BOOL;(*误差刷新标志*)
	axFlag_Refresh_H: ARRAY [1..MAX_UNIT_NUM] OF BOOL;(*误差刷新标志*)
	axFlag_Check_V: ARRAY [1..MAX_UNIT_NUM] OF BOOL;(*误差校验位*)
	axFlag_Check_H: ARRAY [1..MAX_UNIT_NUM] OF BOOL;(*误差校验位*)
	axFlag_PreRefresh_V: ARRAY [1..MAX_UNIT_NUM] OF BOOL;(*误差有效性*)
	axFlag_PreRefresh_H: ARRAY [1..MAX_UNIT_NUM] OF BOOL;(*误差有效性*)
*)	afbKS_FB_PickOutFakePoint_V: ARRAY [1..MAX_UNIT_NUM] OF KS_FB_PickOutFakePoint;(*误差飞点处理*)
	afbKS_FB_PickOutFakePoint_H: ARRAY [1..MAX_UNIT_NUM] OF KS_FB_PickOutFakePoint;
	afbKS_FB_AverageErr_Arc_V: ARRAY [1..MAX_UNIT_NUM] OF KS_FB_AverageErr_Arc;(*误差平均处理*)
	afbKS_FB_AverageErr_Arc_H: ARRAY [1..MAX_UNIT_NUM] OF KS_FB_AverageErr_Arc;
	axFakePoint_V: ARRAY [1..MAX_UNIT_NUM] OF BOOL := [MAX_UNIT_NUM(FALSE)];
	axFakePoint_H: ARRAY [1..MAX_UNIT_NUM] OF BOOL := [MAX_UNIT_NUM(FALSE)];

	aiError_V_Res: ARRAY [1..MAX_UNIT_NUM] OF INT := [MAX_UNIT_NUM(0)];(*处理完成后的纵向误差列表*)
	aiError_H_Res: ARRAY [1..MAX_UNIT_NUM] OF INT := [MAX_UNIT_NUM(0)];(*处理完成后的横向误差列表*)
	abyIndex_V_Pre: ARRAY [1..MAX_UNIT_NUM] OF BYTE := [MAX_UNIT_NUM(0)];(*处理完成后的索引*)
	abyIndex_H_Pre: ARRAY [1..MAX_UNIT_NUM] OF BYTE := [MAX_UNIT_NUM(0)];(*处理完成后的索引*)

	iUnitNR: INT;
	iStationId: INT;
	dwOFST2: DWORD;

	iRtn: INT;
	stStProtocol_PDU_Up_Rd: StParam_PDU_Up;
	pstStCMD_F05_: POINTER TO StPdu_Up_05;
	pbyTemp: POINTER TO BYTE;
	wCHK_Up_Calc: WORD;
	dwCheckSumVal: DWORD;
(*	abyBuf_PduCmd_rcv: ARRAY [1..MAX_PDU_CMD_BYTES_UP] OF BYTE; (* 2021.12.4.163129/hdp/读取 *)*)
(*	xtest: BOOL;*)
	aiResult_VFollowpre_1stDerivate: ARRAY [1..MAX_UNIT_NUM] OF INT := [MAX_UNIT_NUM(0)];

	(*统一注释0916+alTime: ARRAY [1..10] OF LTIME;*)
	abyBuf_PduCmd_rcv_All: ARRAY [1..1000] OF BYTE;

	(*start___@2026.5.10.135832/han.dp
	视觉误差相关的补充变量*)
	adwErrMix_RdVision: ARRAY [1..MAX_UNIT_NUM] OF DWORD := [0];(*来自视觉的复合误差*)
	aiRtnMatrix: ARRAY [1..MAX_UNIT_NUM,1..2] OF INT := [0];(*处理误差解析的返回值矩阵*)
	aiErr_v_pure: ARRAY [1..MAX_UNIT_NUM] OF INT := [0];(*纵向实际误差/从金刚传来/未处理物理坐标系*)
	aiErr_h_pure: ARRAY [1..MAX_UNIT_NUM] OF INT := [0];(*横向实际误差/从金刚传来/未处理物理坐标系*)
(*	adwERR_VisionGave: ARRAY [1..MAX_UNIT_NUM] OF DWORD := [0];(*纵横向误差在一起*)*)

	axFlag_valid_v_tmp: ARRAY [1..MAX_UNIT_NUM] OF BOOL := [MAX_UNIT_NUM(FALSE)];(*纵向有效标志*)
	axFlag_update_v_tmp: ARRAY [1..MAX_UNIT_NUM] OF BOOL := [MAX_UNIT_NUM(FALSE)];(*纵向更新标志*)
	axFlag_update_v_rec: ARRAY [1..MAX_UNIT_NUM] OF BOOL := [MAX_UNIT_NUM(FALSE)];(*纵向上次更新标志*)
	axFlag_bitchk_v_tmp: ARRAY [1..MAX_UNIT_NUM] OF BOOL := [MAX_UNIT_NUM(FALSE)];(*纵向校验位*)

	axFlag_valid_h_tmp: ARRAY [1..MAX_UNIT_NUM] OF BOOL := [MAX_UNIT_NUM(FALSE)];(*横向有效标志*)
	axFlag_update_h_tmp: ARRAY [1..MAX_UNIT_NUM] OF BOOL := [MAX_UNIT_NUM(FALSE)];(*横向更新标志*)
	axFlag_update_h_rec: ARRAY [1..MAX_UNIT_NUM] OF BOOL := [MAX_UNIT_NUM(FALSE)];(*横向上次更新标志*)
	axFlag_bitchk_h_tmp: ARRAY [1..MAX_UNIT_NUM] OF BOOL := [MAX_UNIT_NUM(FALSE)];(*横向校验位*)

	pawErr_tmp: POINTER TO ARRAY [1..2] OF WORD := 0;
	(*___end@2026.5.10.135850*)

	stSystimeDelta,stSystimeStart,stSystimeEnd:SYSTIME;(*获取us时间差*)
	abyVisionErrIdx_V: ARRAY [1..MAX_UNIT_NUM] OF BYTE := [MAX_UNIT_NUM(0)];(*视觉误差索引-纵向*)
	abyVisionErrIdx_H: ARRAY [1..MAX_UNIT_NUM] OF BYTE := [MAX_UNIT_NUM(0)];(*视觉误差索引-横向*)

	xDoNothing: BOOL := FALSE;(*什么都不做*)
	xNeedRead_gLinkII_I_Err: BOOL:= FALSE;
	xNeedRead_gLinkII_II_Err: BOOL:= FALSE;
	iRtn_Rd_I: INT;
	iRtn_Rd_II: INT;
	aiError_V_I: ARRAY [1..MAX_UNIT_NUM] OF INT;(*处理完成后的纵向误差列表*)
	aiError_H_I: ARRAY [1..MAX_UNIT_NUM] OF INT;(*处理完成后的横向误差列表*)
	abyIndex_V_I: ARRAY [1..MAX_UNIT_NUM] OF BYTE;(*处理完成后的索引*)
	abyIndex_H_I: ARRAY [1..MAX_UNIT_NUM] OF BYTE;(*处理完成后的索引*)
	aiError_V_II: ARRAY [1..MAX_UNIT_NUM] OF INT;(*处理完成后的纵向误差列表*)
	aiError_H_II: ARRAY [1..MAX_UNIT_NUM] OF INT;(*处理完成后的横向误差列表*)
(*统一注释0916+	abyErrSts_II: ARRAY [1..MAX_UNIT_NUM] OF BYTE;(*处理完成后的纵横向误差状态*)*)
	abyIndex_V_II: ARRAY [1..MAX_UNIT_NUM] OF BYTE;(*处理完成后的索引*)
	abyIndex_H_II: ARRAY [1..MAX_UNIT_NUM] OF BYTE;(*处理完成后的索引*)
(*统一注释0916+	axValid_V_II: ARRAY [1..MAX_UNIT_NUM] OF BOOL;(*误差有效性*)*)
(*统一注释0916+	axValid_H_II: ARRAY [1..MAX_UNIT_NUM] OF BOOL;(*误差有效性*)	*)
	abyErrSts: ARRAY [1..MAX_UNIT_NUM] OF BYTE;(*处理完成后的纵横向误差状态*)
	axValid_V: ARRAY [1..MAX_UNIT_NUM] OF BOOL;(*误差有效性*)
	axValid_H: ARRAY [1..MAX_UNIT_NUM] OF BOOL;(*误差有效性*)
	aiError_V: ARRAY [1..MAX_UNIT_NUM] OF INT;(*处理完成后的纵向误差列表*)
	aiError_H: ARRAY [1..MAX_UNIT_NUM] OF INT;(*处理完成后的横向误差列表*)
	abyIndex_V: ARRAY [1..MAX_UNIT_NUM] OF BYTE;(*处理完成后的索引*)
	abyIndex_H: ARRAY [1..MAX_UNIT_NUM] OF BYTE;(*处理完成后的索引*)
	xChange_GetErrMode: BOOL;
	(*统一注释0916+2026.4.11.150050+*)
	afbKS_FB_AverageErr_Arc_V_Display: ARRAY [1..MAX_UNIT_NUM] OF KS_FB_AverageErr_Arc;(*误差平均处理@界面显示*)
	afbKS_FB_AverageErr_Arc_H_Display: ARRAY [1..MAX_UNIT_NUM] OF KS_FB_AverageErr_Arc;

	aiError_V_Res_Display: ARRAY [1..MAX_UNIT_NUM] OF INT;(*处理完成后的纵向显示误差列表*)
	aiError_H_Res_Display: ARRAY [1..MAX_UNIT_NUM] OF INT;(*处理完成后的横向显示误差列表*)
	//新飞点剔除:每色组纵横各一个独立实例(总开关gc_xUseNewFlyRemove在GCL)|Yang.zj+用于新飞点检测 2026.10.27.105623
	afbKS_FlyRemove_V: ARRAY [1..MAX_UNIT_NUM] OF KS_FlyRemove;
	afbKS_FlyRemove_H: ARRAY [1..MAX_UNIT_NUM] OF KS_FlyRemove;
	aiError_V_Fly: ARRAY [1..MAX_UNIT_NUM] OF INT;(*剔除后送平均的纵向误差*)
	aiError_H_Fly: ARRAY [1..MAX_UNIT_NUM] OF INT;(*剔除后送平均的横向误差*)
	xFlyNewFrame_V: BOOL;(*本周期该色组纵向是否来了新帧(视觉源纵横索引独立变化,分开判定)*)
	xFlyNewFrame_H: BOOL;(*本周期该色组横向是否来了新帧*)
	xFlyReset: BOOL;(*该色组剔除器复位请求*)
	aiFlyMarkModePre: ARRAY [1..MAX_UNIT_NUM] OF INT;(*上次色标排列模式*)
	abyFlySignalPre: ARRAY [1..MAX_UNIT_NUM] OF BYTE;(*上次RGB信号通道*)
	axFlyHorEnPre: ARRAY [1..MAX_UNIT_NUM] OF BOOL;(*上次横向开关*)
	abyFlyGetErrModePre: ARRAY [1..MAX_UNIT_NUM] OF BYTE;(*上次误差源模式,月光宝盒/金刚切换时复位*)
	axFlyRollPre: ARRAY [1..MAX_UNIT_NUM] OF BOOL;(*上次压辊输出位(g_astStIOMap_Axis_FE[iN].o_xRel_Press,合压继电器原始输出),压下/抬起沿都触发剔除器复位|Yang.zj+ 2026.10.27.210459*)

END_VAR
{IMPLEMENTATION}
SysTimeGetUs(stSystimeStart);(*2026.5.24.152052/han.dp/获取开始时间*)

(*revision by han.dp@2026.5.10.134238*)
o_xEno:= i_xEn;
o_iErNo:= 0;
IF i_xEn THEN
	xChange_GetErrMode:= FALSE;
	FOR iN:=1 TO i_iUnitMax BY 1 DO
		IF abyGetErrMode_Ref[iN]<>i_abyGetErrMode[iN] THEN
			xChange_GetErrMode:= TRUE;
		END_IF
		abyGetErrMode_Ref[iN]:= i_abyGetErrMode[iN];
	END_FOR

	IF xChange_GetErrMode OR
		dwKSMatrixMark_Ref<>i_dwKSMatrixMark THEN
		dwKSMatrixMark_Ref:= i_dwKSMatrixMark;
		IF xInitialized_Ref_KSMatrixMark THEN
			xInitialized_Ref_KSMatrixMark:= FALSE;
		END_IF
	END_IF

	IF NOT xInitialized_Ref_KSMatrixMark THEN
		xInitialized_Ref_KSMatrixMark:= TRUE;

		FOR iN:=1 TO MAX_UNIT_NUM BY 1 DO
			aiRef_KSMatrixMark[iN,1]:= aiRef_KSMatrixMark[iN,2]:= 0;
		END_FOR
		(*生成aiRef_KSMatrixMark*)
		wKSMatrixMark_Hword:= DWORD_TO_WORD(SHR(dwKSMatrixMark_Ref,16) AND 16#FFFF);
		wKSMatrixMark_Lword:= DWORD_TO_WORD(dwKSMatrixMark_Ref AND 16#FFFF);
		IF wKSMatrixMark_Hword=wKSMatrixMark_Lword AND
			wKSMatrixMark_Lword<>0 THEN
			;
		ELSE
			wKSMatrixMark_Hword:= wKSMatrixMark_Lword:= 400;(*默认按1mm直径/1mm间距*)
		END_IF

		(*2026.5.27.100608/han.dp
		*反装顺序和正装逆序/相机成图是一致的
		*按成像后的参考点预置各个色组的0坐标
		*)
		FOR iN:=2 TO 8 BY 1 DO
			IF ((NOT abyGetErrMode_Ref[iN].4) AND abyGetErrMode_Ref[iN].5) OR(*相机正向安装+逆序*)
				(abyGetErrMode_Ref[iN].4 AND (NOT abyGetErrMode_Ref[iN].5)) THEN(*相机反向安装+顺序*)
				IF iN=2 THEN
					aiRef_KSMatrixMark[2,1]:= 0;
					aiRef_KSMatrixMark[2,2]:= WORD_TO_INT(wKSMatrixMark_Hword/2)*(-1);
				END_IF
				IF iN=3 THEN
					aiRef_KSMatrixMark[3,1]:= WORD_TO_INT(wKSMatrixMark_Hword/2)*(-1);
					aiRef_KSMatrixMark[3,2]:= WORD_TO_INT(wKSMatrixMark_Hword/2)*(-1);
				END_IF
				IF iN=4 THEN
					aiRef_KSMatrixMark[4,1]:= WORD_TO_INT(wKSMatrixMark_Hword/2);
					aiRef_KSMatrixMark[4,2]:= 0;
				END_IF
				IF iN=5 THEN
					aiRef_KSMatrixMark[5,1]:= 0;
					aiRef_KSMatrixMark[5,2]:= 0;
				END_IF
				IF iN=6 THEN
					aiRef_KSMatrixMark[6,1]:= WORD_TO_INT(wKSMatrixMark_Hword/2)*(-1);
					aiRef_KSMatrixMark[6,2]:= 0;
				END_IF
				IF iN=7 THEN
					aiRef_KSMatrixMark[7,1]:= WORD_TO_INT(wKSMatrixMark_Hword/2);
					aiRef_KSMatrixMark[7,2]:= WORD_TO_INT(wKSMatrixMark_Hword/2);
				END_IF
				IF iN=8 THEN
					aiRef_KSMatrixMark[8,1]:= 0;
					aiRef_KSMatrixMark[8,2]:= WORD_TO_INT(wKSMatrixMark_Hword/2);
				END_IF
			ELSE
				IF iN=2 THEN
					aiRef_KSMatrixMark[2,1]:= 0;
					aiRef_KSMatrixMark[2,2]:= WORD_TO_INT(wKSMatrixMark_Hword/2);
				END_IF

				IF iN=3 THEN
					aiRef_KSMatrixMark[3,1]:= WORD_TO_INT(wKSMatrixMark_Hword/2);
					aiRef_KSMatrixMark[3,2]:= WORD_TO_INT(wKSMatrixMark_Hword/2);
				END_IF

				IF iN=4 THEN
					aiRef_KSMatrixMark[4,1]:= WORD_TO_INT(wKSMatrixMark_Hword/2)*(-1);
					aiRef_KSMatrixMark[4,2]:= 0;
				END_IF

				IF iN=5 THEN
					aiRef_KSMatrixMark[5,1]:= 0;
					aiRef_KSMatrixMark[5,2]:= 0;
				END_IF

				IF iN=6 THEN
					aiRef_KSMatrixMark[6,1]:= WORD_TO_INT(wKSMatrixMark_Hword/2);
					aiRef_KSMatrixMark[6,2]:= 0;
				END_IF

				IF iN=7 THEN
					aiRef_KSMatrixMark[7,1]:= WORD_TO_INT(wKSMatrixMark_Hword/2)*(-1);
					aiRef_KSMatrixMark[7,2]:= WORD_TO_INT(wKSMatrixMark_Hword/2)*(-1);
				END_IF

				IF iN=8 THEN
					aiRef_KSMatrixMark[8,1]:= 0;
					aiRef_KSMatrixMark[8,2]:= WORD_TO_INT(wKSMatrixMark_Hword/2)*(-1);
				END_IF
			END_IF
		END_FOR
	END_IF

(*统一注释0916+重新整理一下逻辑*)
	xNeedRead_gLinkII_I_Err:=FALSE;
	xNeedRead_gLinkII_II_Err:= FALSE;
	IF (i_iUnitMax>0 AND i_iUnitMax<=MAX_UNIT_NUM) THEN

		FOR iN:= 1 TO i_iUnitMax BY 1 DO
			IF i_abyGetErrMode[iN].0 THEN(*统一注释0916+有一个色组打开了读取月光宝盒误差*)
				xNeedRead_gLinkII_I_Err:= TRUE;
			END_IF
		END_FOR
		FOR iN:= 1 TO i_iUnitMax BY 1 DO
			IF i_abyGetErrMode[iN].1 THEN(*统一注释0916+有一个色组打开了读取金刚误差*)
				xNeedRead_gLinkII_II_Err:= TRUE;
			END_IF
		END_FOR
	END_IF
(*统一注释0916+读取地址*)
iRtn_Rd_I:= -1;
iRtn_Rd_II:= -1;
	IF (NOT xNeedRead_gLinkII_II_Err) AND (NOT xNeedRead_gLinkII_I_Err) THEN(*统一注释0916+2026.5.30.090808都没有默认读一下一套网内容*)
		iRtn_Rd_I :=
			GTN_RN_UserPCRdLocalFPGA(
				1(*cardIndex*),
				1(*busIndex*),
				0(*stationId*),
				ADR(abyBuf_PduCmd_rcv_All)(*pData*),
				0(*startAddr*),
				KS_GetNumOfDwordUsed(INT_TO_DWORD(i_iUnitMax)*MAX_PDU_CMD_BYTES_DN)(*dwordNum*));

	ELSE
		IF xNeedRead_gLinkII_I_Err THEN
			iRtn_Rd_I :=
				GTN_RN_UserPCRdLocalFPGA(
					1(*cardIndex*),
					1(*busIndex*),
					0(*stationId*),
					ADR(abyBuf_PduCmd_rcv_All)(*pData*),
					0(*startAddr*),
					KS_GetNumOfDwordUsed(INT_TO_DWORD(i_iUnitMax)*MAX_PDU_CMD_BYTES_DN)(*dwordNum*));

		END_IF
		IF xNeedRead_gLinkII_II_Err THEN
			iRtn_Rd_II:=
				GTN_RN_GetVisualControllerValue(
					1(*cardIndex*),
					2(*busIndex*),
					ADR(adwErrMix_RdVision)(*pData*),
					MAX_UNIT_NUM(*dwordNum*));
		END_IF
	END_IF
(*统一注释0916+地址读取完成，把读到的内容处理一遍	*)
	IF iRtn_Rd_I=0 THEN(*统一注释0916+这里先这样处理吧？一套网的协议解析一下*)
		FOR iN:=1 TO i_iUnitMax BY 1 DO
			iUnitNR:= iN;(*通讯轴号也需要根据后续系统配置处理*)
			iStationId:= g_stStSysParam.stStSysParam_UnSave.aiStationList_UnitController[iN];(*统一注释0916+g_abyStationList_CommKSCR[iN];(*站号*)*)
			IF KS_IsValidStationNR(iStationId) THEN(*站号有效*)
				dwOFST2 := MAX_PDU_CMD_BYTES_DN*(iUnitNR-1);(*偏移量*)
				SysMemCpy(
					ADR(stStProtocol_PDU_Up_Rd),
					ADR(abyBuf_PduCmd_rcv_All)+dwOFST2,
					SIZEOF(stStProtocol_PDU_Up_Rd));

				(*2026.5.10.143526/han.dp/从16#5号命令解析内部移出来*)
				aiError_V_I[iN]:= stStProtocol_PDU_Up_Rd.iErr_V_Raw;
				aiError_H_I[iN]:= stStProtocol_PDU_Up_Rd.iErr_H_Raw;
				abyIndex_V_I[iN]:= stStProtocol_PDU_Up_Rd.byIDX_V;
				abyIndex_H_I[iN]:= stStProtocol_PDU_Up_Rd.byIDX_H;

				(*2026.10.24.180455+*)
				o_astStErrParam_Use[iN].uiFSampleCounter:=stStProtocol_PDU_Up_Rd.uiFSampleCounter;
				i_pstStSysParam^.astStUnitParam_UnSave[iN].uiFSampleCounter:=stStProtocol_PDU_Up_Rd.uiFSampleCounter;

				(*2026.09.15.134645//xi.hy//增加月光宝盒Pro另一路误差的保存*)
				g_aiError_V_Other[iN]:=stStProtocol_PDU_Up_Rd.iErr_V_Raw_1;
				g_aiError_H_Other[iN]:=stStProtocol_PDU_Up_Rd.iErr_H_Raw_1;

				(*如果附加的报文是命令/如下便是解析过程*)
				pbyTemp:= ADR(stStProtocol_PDU_Up_Rd.byPkgId);
				wCHK_Up_Calc:= KS_CRC(pbyTemp, 46, ADR(dwCheckSumVal));(*46=byPkgId+abyPayLoad的长度*)
				IF wCHK_Up_Calc=stStProtocol_PDU_Up_Rd.wCHK THEN(*CRC校验OK*)
					CASE stStProtocol_PDU_Up_Rd.byPkgId OF
					16#5:(*command of 'StPdu_Up_05'*)
						pstStCMD_F05_:= ADR(stStProtocol_PDU_Up_Rd.abyPayload);
						IF pstStCMD_F05_<>0 THEN
							o_astStErrParam_Use[iN].iResult_VFollowpre_1stDerivate:= pstStCMD_F05_^.iResult_VFollowpre_1stDerivate;
							aiResult_VFollowpre_1stDerivate[iN]:= pstStCMD_F05_^.iResult_VFollowpre_1stDerivate;
							o_astStErrParam_Use[iN].uiBaseUse_t1:= pstStCMD_F05_^.uiBaseUse_t1;
							o_astStErrParam_Use[iN].uiBaseUse_t2:= pstStCMD_F05_^.uiBaseUse_t2;
							o_astStErrParam_Use[iN].uiPeakValue_t1:= pstStCMD_F05_^.uiPeakValue_t1;
							o_astStErrParam_Use[iN].uiPeakValue_t2:= pstStCMD_F05_^.uiPeakValue_t2;
						(*统一注释0916+2026.5.9.110642	*)
							i_pstStSysParam^.astStRSV_UnitParam_UnSave[iN].iCurLabelPos:= pstStCMD_F05_^.iCurLabelPos;(*本色三角标位置，点数*)
							i_pstStSysParam^.astStRSV_UnitParam_UnSave[iN].iPreLabelPos:= pstStCMD_F05_^.iPreLabelPos;(*前色三角标位置，点数*)
							i_pstStSysParam^.astStRSV_UnitParam_UnSave[iN].byFlag_CommFromSlave:= pstStCMD_F05_^.byFlag_CommFromSlave;(*bit0 xFlag_FindFirstSuccess;bit1 xFlag_FindPreSuccess*)
							i_pstStSysParam^.astStRSV_UnitParam_UnSave[iN].xFlag_FindFirstSuccess:= i_pstStSysParam^.astStRSV_UnitParam_UnSave[iN].byFlag_CommFromSlave.0;
							i_pstStSysParam^.astStRSV_UnitParam_UnSave[iN].xFlag_FindPreSuccess:= i_pstStSysParam^.astStRSV_UnitParam_UnSave[iN].byFlag_CommFromSlave.1;
							i_pstStSysParam^.astStRSV_UnitParam_UnSave[iN].byDetectedSignalCount:= pstStCMD_F05_^.byDetectedSignalCount;(*当前检测到色标个数*)
							i_pstStSysParam^.astStRSV_UnitParam_UnSave[iN].byMarkStep:= pstStCMD_F05_^.byMarkStep;(*当前全自动套印步骤*)
							i_pstStSysParam^.astStRSV_UnitParam_UnSave[iN].rGateSignalWidth_R:= BYTE_TO_REAL (pstStCMD_F05_^.byWidthRS) /10.0;(*粗采样计算波形宽度*)

						END_IF
					ELSE;
					END_CASE
				END_IF
			END_IF
		END_FOR(*end?'FOR iN:=1 TO i_iUnitMax BY 1 DO'*)
	ELSE;
	END_IF

	IF iRtn_Rd_II=0 THEN
		(*开始逐色组处理读取的内容*)
		FOR iN:=2 TO i_iUnitMax BY 1 DO(*2026.5.24.212501/han.dp/套色误差是从2色开始的*)
			pawErr_tmp:= ADR(adwErrMix_RdVision[iN-1]);

			(*纵向误差*)
			aiRtnMatrix[iN,1]:=
			KS_UnPack_VisionERR(
				pawErr_tmp^[1],(*2026.5.27.102650/han.dp/按原理梳理/第1个数值是相机检测的X距离/顺时针90度旋转成了Y*)
				ADR(axFlag_valid_v_tmp[iN]),
				ADR(axFlag_update_v_tmp[iN]),
				ADR(axFlag_bitchk_v_tmp[iN]),
				ADR(aiERR_v_pure[iN]));
			IF aiRtnMatrix[iN,1]=0 THEN(*转换ok*)
				IF axFlag_update_v_tmp[iN]<>axFlag_update_v_rec[iN] THEN(*误差更新了*)
					o_astStErrParam_Use[iN].uiV_cam_raw:= pawErr_tmp^[1];
					IF axFlag_valid_v_tmp[iN] THEN(*误差有效*)
						aiError_V_II[iN]:= -aiERR_v_pure[iN] - aiRef_KSMatrixMark[iN,2];(*2026.5.27.110642/han.dp/方向修订*)
					ELSE(*误差无效*)
						aiError_V_II[iN]:= gc_iValueReferToLost;
					END_IF
					abyIndex_V_II[iN]:= abyIndex_V_II[iN]+1;
				END_IF
				axFlag_update_v_rec[iN]:= axFlag_update_v_tmp[iN];
			END_IF

			(*横向误差*)
			aiRtnMatrix[iN,2]:=
			KS_UnPack_VisionERR(
				pawErr_tmp^[2],
				ADR(axFlag_valid_h_tmp[iN]),
				ADR(axFlag_update_h_tmp[iN]),
				ADR(axFlag_bitchk_h_tmp[iN]),
				ADR(aiERR_h_pure[iN]));
			IF aiRtnMatrix[iN,2]=0 THEN(*转换ok*)
				IF axFlag_update_h_tmp[iN]<>axFlag_update_h_rec[iN] THEN(*误差更新了*)
					axFlag_update_h_rec[iN]:= axFlag_update_h_tmp[iN];
					o_astStErrParam_Use[iN].uiH_cam_raw:= pawErr_tmp^[2];
					IF axFlag_valid_h_tmp[iN] THEN(*误差有效*)
						aiError_H_II[iN]:= -aiERR_h_pure[iN] - aiRef_KSMatrixMark[iN,1];(*2026.5.27.132504/han.dp/修订方向*)
					ELSE(*误差无效*)
						aiError_H_II[iN]:= gc_iValueReferToLost;
					END_IF
					abyIndex_H_II[iN]:= abyIndex_H_II[iN]+1;
				END_IF
			END_IF
		END_FOR
	ELSE;
	END_IF
	(*统一注释0916+2026.5.30.094300*)
	FOR iN:=1 TO i_iUnitMax BY 1 DO
		IF i_abyGetErrMode[iN].1 AND i_abyGetErrMode[iN].7 THEN(*统一注释0916+指定了金刚并且打开了金刚误差调整*)
			abyIndex_V[iN]:= abyIndex_V_II[iN];
			abyIndex_H[iN]:= abyIndex_H_II[iN];
			aiError_V[iN]:= aiError_V_II[iN];
			aiError_H[iN]:= aiError_H_II[iN];
		ELSE(*统一注释0916+其他全部按月光宝盒误差处理吧*)
			abyIndex_V[iN]:= abyIndex_V_I[iN];
			abyIndex_H[iN]:= abyIndex_H_I[iN];
			aiError_V[iN]:= aiError_V_I[iN];
			aiError_H[iN]:= aiError_H_I[iN];
		END_IF

(*统一注释0916+加保存吧2026.5.30.095819*)
		o_astStErrParam_Use[iN].iV_cam_pure:= aiError_V_II[iN];
		o_astStErrParam_Use[iN].iH_cam_pure:= aiError_H_II[iN];
		o_astStErrParam_Use[iN].iErr_V_I_:= aiError_V_I[iN];
		o_astStErrParam_Use[iN].iErr_H_I_:= aiError_H_I[iN];
(*统一注释0916+到这里误差已经有了，处理各种标志*)
		(*新飞点剔除:误差平均之前对原始逐帧误差剔除,飞点/暂缓用锁存值(上一好值)替换,必须先剔除再平均,否则飞点被N幅平均稀释后可能低于门限漏掉*
		 *本版纵/横索引可能独立变化(金刚视觉源),故按各自索引变化判定新帧;总开关gc_xUseNewFlyRemove在GCL,置FALSE并重编译即回退旧逻辑*
		 *飞点/暂缓帧置axFakePoint_V/H(byErrSts.2/6),阶跃(真实变化)不置位|Yang.zj+用于新飞点检测 2026.10.27.105623*)
		IF gc_xUseNewFlyRemove THEN
			xFlyNewFrame_V:= (abyIndex_V_Pre[iN]<>abyIndex_V[iN]);
			xFlyNewFrame_H:= (abyIndex_H_Pre[iN]<>abyIndex_H[iN]);
			(*工况切换检测:色标排列模式/RGB信号通道/横向开关/误差源模式任一变化,该色组剔除器可信历史不可信,复位重新暖机*)
			xFlyReset:= FALSE;
			IF i_pstStSysParam<>0 THEN
				IF (aiFlyMarkModePre[iN]<>i_pstStSysParam^.astStUnitParam_Save[iN].iMarkArrangeMode)
					OR (abyFlySignalPre[iN]<>i_pstStSysParam^.astStUnitParam_Save[iN].bySignalSelect)
					OR (axFlyHorEnPre[iN]<>i_pstStSysParam^.astStUnitParam_Save[iN].dwFlag_Ctl.0)
					OR (abyFlyGetErrModePre[iN]<>i_abyGetErrMode[iN])
					OR (axFlyRollPre[iN]<>g_astStIOMap_Axis_FE[iN].o_xRel_Press) THEN(*压辊沿:合压/抬起双向变化都复位——停机/急停同样引起压辊变化,一并覆盖;安静期旧σ与历史对压辊后快速爬坡完全不适用,不复位会陷入"确认→观察失败"两帧循环,输出冻结(实测4U开机压辊冻结15帧/约47秒)|Yang.zj+ 2026.10.27.210459*)
					aiFlyMarkModePre[iN]:= i_pstStSysParam^.astStUnitParam_Save[iN].iMarkArrangeMode;
					abyFlySignalPre[iN]:= i_pstStSysParam^.astStUnitParam_Save[iN].bySignalSelect;
					axFlyHorEnPre[iN]:= i_pstStSysParam^.astStUnitParam_Save[iN].dwFlag_Ctl.0;
					abyFlyGetErrModePre[iN]:= i_abyGetErrMode[iN];
					axFlyRollPre[iN]:= g_astStIOMap_Axis_FE[iN].o_xRel_Press;
					xFlyReset:= TRUE;
				END_IF
			END_IF
			afbKS_FlyRemove_V[iN](
				i_iErr:= aiError_V[iN],
				i_xErrValid:= xFlyNewFrame_V AND (aiError_V[iN]<>gc_iValueReferToLost),
				i_xLost:= xFlyNewFrame_V AND (aiError_V[iN]=gc_iValueReferToLost),
				i_xReset:= xFlyReset,
				o_iErrResult=> aiError_V_Fly[iN],
				o_xFake=> axFakePoint_V[iN]);
			afbKS_FlyRemove_H[iN](
				i_iErr:= aiError_H[iN],
				i_xErrValid:= xFlyNewFrame_H AND (aiError_H[iN]<>gc_iValueReferToLost),
				i_xLost:= xFlyNewFrame_H AND (aiError_H[iN]=gc_iValueReferToLost),
				i_xReset:= xFlyReset,
				o_iErrResult=> aiError_H_Fly[iN],
				o_xFake=> axFakePoint_H[iN]);
		ELSE
			aiError_V_Fly[iN]:= aiError_V[iN];(*旧路径:不剔除,原值送平均*)
			aiError_H_Fly[iN]:= aiError_H[iN];
		END_IF
		IF abyIndex_V_Pre[iN]<>abyIndex_V[iN] OR abyIndex_H_Pre[iN]<>abyIndex_H[iN] THEN
			abyErrSts[iN]:= 0;
			axValid_V[iN]:= FALSE;
			axValid_H[iN]:= FALSE;

			IF aiError_V[iN]=gc_iValueReferToLost THEN
				abyErrSts[iN].1:= TRUE;(*纵向丢失*)
			ELSE
				axValid_V[iN]:= TRUE;
			END_IF

			IF aiError_H[iN]=gc_iValueReferToLost THEN
				abyErrSts[iN].5:= TRUE;(*横向丢失*)
			ELSE
				axValid_H[iN]:= TRUE;
			END_IF

			o_astStErrParam_Use[iN].byIDX_V:= abyIndex_V[iN];
			o_astStErrParam_Use[iN].byIDX_H:= abyIndex_H[iN];

			(*误差平均-纵向*)
			afbKS_FB_AverageErr_Arc_V[iN](
				i_xEn:= TRUE,
				i_iErr:= aiError_V_Fly[iN],(*新飞点:喂剔除后的值|Yang.zj+用于新飞点检测 2026.10.27.105623*)
				i_xErrValid:= axValid_V[iN],(*2025.01.03.110017*)
				i_byAverageNum:= i_abyAverageNum_V[iN],
				o_iErrResult=>aiError_V_Res[iN]);

			IF NOT gc_xUseNewFlyRemove THEN(*旧飞点判断:新算法启用时整块跳过|Yang.zj+用于新飞点检测 2026.10.27.105623*)
			(*飞点剔除-纵向*)
			axFakePoint_V[iN]:= FALSE;
			afbKS_FB_PickOutFakePoint_V[iN](
				i_xIsValidError:= axValid_V[iN],
				i_iError_0_01mm:= aiError_V_Res[iN],
				i_iVariationBaseValue:= 50,(*2025.01.03.110017*)
				i_iBoundaryError_0_01mm:= 20,
				i_iErrorLevel_0_01mm:= 25,
				i_iVariationVariationMin:= 5,
				i_iVariationVariationMax:= 50,
				o_xFakeIsConfirmed=> axFakePoint_V[iN]);
			END_IF

			(*误差平均-横向*)
			afbKS_FB_AverageErr_Arc_H[iN](
				i_xEn:= TRUE,
				i_iErr:= aiError_H_Fly[iN],(*新飞点:喂剔除后的值|Yang.zj+用于新飞点检测 2026.10.27.105623*)
				i_xErrValid:= axValid_H[iN],(*2025.01.03.110017*)
				i_byAverageNum:= i_abyAverageNum_H[iN],
				o_iErrResult=>aiError_H_Res[iN]);

			IF NOT gc_xUseNewFlyRemove THEN(*旧飞点判断:新算法启用时整块跳过|Yang.zj+用于新飞点检测 2026.10.27.105623*)
			(*飞点剔除-横向*)
			axFakePoint_H[iN]:= FALSE;
			afbKS_FB_PickOutFakePoint_H[iN](
				i_xIsValidError:= axValid_H[iN],
				i_iError_0_01mm:= aiError_H_Res[iN],
				i_iVariationBaseValue:= 50,
				i_iBoundaryError_0_01mm:= 20,
				i_iErrorLevel_0_01mm:= 25,
				i_iVariationVariationMin:= 5,
				i_iVariationVariationMax:= 50,
				o_xFakeIsConfirmed=> axFakePoint_H[iN]);
			END_IF
			(*统一注释0916+显示平均@2026.4.11.150119+	*)
			afbKS_FB_AverageErr_Arc_V_Display[iN](
				i_xEn:= TRUE,
				i_iErr:= aiError_V_Fly[iN],(*新飞点:喂剔除后的值|Yang.zj+用于新飞点检测 2026.10.27.105623*)
				i_xErrValid:= axValid_V[iN],(*2025.01.03.110017*)
				i_byAverageNum:= i_abyAverageNum_V_Display[iN],
				o_iErrResult=>aiError_V_Res_Display[iN]);

			afbKS_FB_AverageErr_Arc_H_Display[iN](
				i_xEn:= TRUE,
				i_iErr:= aiError_H_Fly[iN],(*新飞点:喂剔除后的值|Yang.zj+用于新飞点检测 2026.10.27.105623*)
				i_xErrValid:= axValid_H[iN],(*2025.01.03.110017*)
				i_byAverageNum:= i_abyAverageNum_H_Display[iN],
				o_iErrResult=>aiError_H_Res_Display[iN]);

		END_IF
		(*到这里误差的飞点和平均都处理完了，该处理其他东西了*)
		o_astStErrParam_Use[iN].iErr_V_Unprocessed:= aiError_V[iN];(*原始误差*)
		o_astStErrParam_Use[iN].iErr_H_Unprocessed:= aiError_H[iN];

		o_astStErrParam_Use[iN].byErrSts:= 0;
		o_astStErrParam_Use[iN].byErrSts:= abyErrSts[iN];(*现在的状态*)

(*统一注释0916+2026.5.9.110835处理一下显示平均相关			*)
		IF NOT o_astStErrParam_Use[iN].byErrSts.1 THEN(*纵向未丢失*)
			o_astStErrParam_Use[iN].iErr_V:= aiError_V_Res[iN]-i_aiAdjust_V[iN];
			(*统一注释0916+2026.4.11.150603+*)
			o_astStErrParam_Use[iN].iErr_V_Display:= aiError_V_Res_Display[iN]-i_aiAdjust_V[iN];
			IF axFakePoint_V[iN] THEN(*飞点*)
				o_astStErrParam_Use[iN].byErrSts.2:= TRUE;
			END_IF
			(*报警标志检查*)
			IF ABS(o_astStErrParam_Use[iN].iErr_V_Display)>ABS(i_aiAlarm_V[iN]) THEN
				o_astStErrParam_Use[iN].byErrSts.0:= TRUE;
			END_IF
		ELSE
			o_astStErrParam_Use[iN].iErr_V:= gc_iValueReferToLost;
			o_astStErrParam_Use[iN].iErr_V_Display:= gc_iValueReferToLost;
		END_IF
		IF NOT o_astStErrParam_Use[iN].byErrSts.5 THEN(*横向未丢失*)
			o_astStErrParam_Use[iN].iErr_H:= aiError_H_Res[iN]-i_aiAdjust_H[iN];(*处理完的误差-修正量*)
			(*统一注释0916+2026.4.11.150603+*)
			o_astStErrParam_Use[iN].iErr_H_Display:= aiError_H_Res_Display[iN]-i_aiAdjust_H[iN];
			IF axFakePoint_H[iN] THEN(*飞点*)
				o_astStErrParam_Use[iN].byErrSts.6:= TRUE;
			END_IF
			(*报警标志检查*)
			IF ABS(o_astStErrParam_Use[iN].iErr_H_Display)>ABS(i_aiAlarm_H[iN]) THEN
				o_astStErrParam_Use[iN].byErrSts.4:= TRUE;
			END_IF
		ELSE
			o_astStErrParam_Use[iN].iErr_H:= gc_iValueReferToLost;
			(*统一注释0916+2026.4.11.150603+*)
			o_astStErrParam_Use[iN].iErr_H_Display:= gc_iValueReferToLost;
		END_IF
		abyIndex_V_Pre[iN]:= abyIndex_V[iN];
		abyIndex_H_Pre[iN]:= abyIndex_H[iN];
	END_FOR
END_IF

SysTimeGetUs(stSystimeEnd);(*2026.5.24.152052/han.dp/获取结束时间*)
o_stSystimeElapsed:= stSystimeEnd-stSystimeStart;(*耗时/单位us*)

(* ---- KS_FB_PickOutFakePoint.st ---- *)
(*@CES
Name=KS_FB_PickOutFakePoint
Type=FunctionBlock
TypeGuid=6f9dac99-8de1-4efc-8465-68ac443b7d08
Guid=a2f1e1a0-e198-4123-93c4-db1d31fdab22
HasDeclaration=True
HasImplementation=True
*)
{DECLARATION}
FUNCTION_BLOCK KS_FB_PickOutFakePoint
VAR_INPUT
	i_xIsValidError							: BOOL; (*the error is valid or invalid; TRUE :is valid;*)
	i_iError_0_01mm							: INT; (*error value, unit in 0.01mm*)
	i_iVariationBaseValue					: INT  := 5; (*based variation threshold*)
	i_iBoundaryError_0_01mm					: INT  := 50; (*Boundary error*)
	i_iErrorLevel_0_01mm					: INT  := 25; (*error value per level when up than boundary error.*)
	i_iVariationVariationMin				: INT  := 5; (*minimized variation variation*)
	i_iVariationVariationMax				: INT  := 15; (*maximized variation variation*)
END_VAR
VAR_OUTPUT
	o_xFakeIsConfirmed						: BOOL; (*TRUE :confirm is fake error; FALSE :confirm is normal error*)
END_VAR
VAR
	iN										: INT;
	iUsedVariationMaxThreshold				: INT;
	aiBufferedError							: ARRAY [1..3] OF INT; (*buffered error list*)
	aiVariation								: ARRAY [1..2] OF INT; (*variation*)
	iVariationVariation						: INT; (*variation's variation*)
END_VAR

{IMPLEMENTATION}
IF NOT i_xIsValidError THEN (*invalid error process*)
	o_xFakeIsConfirmed:= TRUE;
	aiBufferedError[1]:= 0;
	aiBufferedError[2]:= 0;
	aiBufferedError[3]:= 0;
ELSE (*valid error process*)
	(*误差变化量的变化量不超出10|2016.10.14.120106_*)
	IF ABS(i_iError_0_01mm)<=i_iBoundaryError_0_01mm THEN (*0.5mm内的误差变化量的变化量不超过5不认为是飞点*)
		iUsedVariationMaxThreshold:= i_iVariationBaseValue;
	ELSE
		iUsedVariationMaxThreshold:= i_iVariationBaseValue+(ABS(i_iError_0_01mm)-i_iBoundaryError_0_01mm)/i_iErrorLevel_0_01mm; (*超过0.5mm的误差,每0.25mm一个档位递增变化量的变化量*)
		IF iUsedVariationMaxThreshold>i_iVariationVariationMax THEN (*upper limit*)
			iUsedVariationMaxThreshold:= i_iVariationVariationMax;
		ELSIF iUsedVariationMaxThreshold<i_iVariationVariationMin THEN (*lower limit*)
			iUsedVariationMaxThreshold:= i_iVariationVariationMin;
		END_IF
	END_IF

	(*存放规则:都是用下标1来记录当前误差|2017.3.31.145925_*)
	(*rolling the buffered error list*)
	FOR iN:=3 TO 2 BY -1 DO
		aiBufferedError[iN]:= aiBufferedError[iN-1];
	END_FOR
	aiBufferedError[1]:= i_iError_0_01mm; (*record the current error to buffered error list*)

	(*calculate error variation*)
	FOR iN:=3 TO 2 BY -1 DO
		aiVariation[iN-1]:= aiBufferedError[iN-1]-aiBufferedError[iN]; (*new - old*)
	END_FOR

	(*calculate error variation variation*)
	iVariationVariation:= aiVariation[1] - aiVariation[2];

	IF ABS(iVariationVariation)>ABS(iUsedVariationMaxThreshold) THEN
		o_xFakeIsConfirmed:= TRUE;
	ELSE
		o_xFakeIsConfirmed:= FALSE;
	END_IF
END_IF

(* ---- KS_FlyRemove.st ---- *)
(*@CES
Name=KS_FlyRemove
Type=FunctionBlock
TypeGuid=6f9dac99-8de1-4efc-8465-68ac443b7d08
Guid=ea8acba0-5633-4be0-8daa-610d8883b0ed
HasDeclaration=True
HasImplementation=True
*)
{DECLARATION}
FUNCTION_BLOCK KS_FlyRemove
VAR_INPUT
	i_iErr			: INT;	(*原始误差|丝*)
	i_xErrValid		: BOOL;	(*TRUE=本帧为有效新帧(喂入剔除);FALSE=不喂*)
	i_xLost			: BOOL;	(*TRUE=本帧为丢失帧(原样上报-32768,不算飞点)*)
	i_xReset		: BOOL;	(*TRUE=复位全部状态(工况切换时给一拍)*)
END_VAR
VAR_OUTPUT
	o_iErrResult	: INT;	(*剔除后输出:好=原值,飞点/暂缓=锁存值,丢失=原值原样*)
	o_byJudge		: BYTE;	(*0首帧 1好 2好(观察) 3飞点 4暂缓 5阶跃 6丢失*)
	o_xFake			: BOOL;	(*本帧输出被替换(飞点/暂缓)=TRUE;阶跃/丢失/好=FALSE*)
END_VAR
VAR
	KS_FLY_TRUST_WIN	: INT	:= 9;	(*趋势窗:Theil-Sen用最近N个可信点*)
	KS_FLY_NOISE_WIN	: INT	:= 31;	(*噪声窗:差分rSigma用最近N个可信值*)
	KS_FLY_DIFF_MIN		: INT	:= 8;	(*差分数不足N不用MAD(防越剔越紧螺旋)*)
	KS_FLY_SIG_PROV		: REAL	:= 2.0;	(*暖机rSigma倍数(尺度自举,量纲无关)*)
	KS_FLY_K			: REAL	:= 5.0;	(*外门槛倍数:T_out=K*rSigma*)
	KS_FLY_RET_FRAC		: REAL	:= 0.5;	(*回归门槛=该比例*外门槛(5rSigma/2.5rSigma)*)
	KS_FLY_STEP_CONFIRM	: INT	:= 2;	(*阶跃确认:连续强超门满N帧判阶跃*)
	KS_FLY_QUAR_N		: INT	:= 1;	(*阶跃确认后的观察帧数*)
	KS_FLY_HOLD_MAX		: INT	:= 3;	(*迟滞带内暂缓上限(暂缓不等于剔除)*)
	KS_FLY_OSC_WIN		: INT	:= 64;	(*振荡自愈:统计近N帧判非好占比*)
	KS_FLY_OSC_IN		: REAL	:= 0.25;	(*振荡模式进入门限*)
	KS_FLY_OSC_OUT		: REAL	:= 0.10;	(*振荡模式退出门限*)
	KS_FLY_MAD_C		: REAL	:= 1.4826;		(*MAD->正态标准差一致性系数*)
	KS_FLY_SQRT2		: REAL	:= 1.414213562;	(*根2:Var(差分)=2*rSigma^2的归一*)
	KS_FLY_EPS			: REAL	:= 1.0E-12;		(*rSigma=0保护*)
	(*状态:逐项对应C版KsFlyRemover结构体*)
	arHistVal	: ARRAY[0..30] OF REAL;		(*可信历史值:只有真实测量进*)
	auiHistIdx	: ARRAY[0..30] OF UDINT;	(*各历史点帧号(内部稠密计数,严格递增)*)
	iHistCnt	: INT;						(*历史点数(<=31)*)
	xStarted	: BOOL;						(*启动态:前2帧无条件采信;阶跃重建不回退此标志*)
	rLatch		: REAL;						(*锁存:最近好值,飞点替换用它;只被好帧更新*)
	xLatchValid	: BOOL;
	rSigma		: REAL;						(*差分MAD的rSigma估计*)
	xSigmaValid	: BOOL;						(*未估出时用暖机rSigma;阶跃只换电平不换噪声*)
	iConsec		: INT;						(*连续强超门计数(阶跃确认用)*)
	iQuar		: INT;						(*阶跃确认后的观察帧余数*)
	iHold		: INT;						(*候选期暂缓计数*)
	abyJudged	: ARRAY[0..63] OF BYTE;		(*近64帧是否判非好(振荡自愈检测用)*)
	iJudgedCnt	: INT;
	arAllDev	: ARRAY[0..15] OF REAL;		(*近16帧|新值-带中心|(含被拒帧,振荡模式估幅用)*)
	iAllDevCnt	: INT;
	xOscOn		: BOOL;						(*振荡模式开关(生效时门放宽到全幅MAD)*)
	udiIdxNext	: UDINT;					(*下一帧帧号(丢失帧不占号)*)
	(*中位数运算暂存区*)
	arSlope		: ARRAY[0..35] OF REAL;		(*Theil-Sen两两斜率(9点36对)*)
	arExt		: ARRAY[0..8] OF REAL;		(*趋势带:外推值/水平值的中位数暂存*)
	arDiff		: ARRAY[0..29] OF REAL;		(*可信历史相邻差分(<=30个)*)
	arDev		: ARRAY[0..15] OF REAL;		(*全幅偏差中位数暂存(振荡模式)*)
	(*工作变量*)
	rX			: REAL;
	rOut		: REAL;
	rA			: REAL;
	rB			: REAL;
	rD			: REAL;
	rS			: REAL;
	rTOut		: REAL;
	rTRet		: REAL;
	rRatio		: REAL;
	rTmp		: REAL;
	rMed		: REAL;
	fV			: REAL;
	fP			: REAL;
	fL			: REAL;
	i			: INT;
	j			: INT;
	n			: INT;
	m			: INT;
	iSum		: INT;
	udiIdx		: UDINT;
	udiDt		: UDINT;
	iBase		: INT;
	byJudge		: BYTE;
	(*为了加 Quantum 去处理稳态的小范围波动不报飞点*)
	arQdq		: ARRAY[0..15] OF REAL;		(*近16个非零相邻差分,数据分辨率quantum用|Yang.zj 2026.10.27+*)
	iQdqCnt		: INT;
	rPval		: REAL;						(*上一有效输入值(含被拒帧,算分辨率用)*)
	xPvalValid	: BOOL;
	udiPidx		: UDINT;					(*上一有效输入帧号(跨丢失段的差分不入分辨率)*)
	rQuantum	: REAL;						(*数据分辨率=近16个非零相邻差分最小值(需>=2个样本)*)
	xQuantumValid	: BOOL;
END_VAR

{IMPLEMENTATION}
(*==================== 复位:清零全部状态(工况切换时) ====================*)
IF i_xReset THEN
	iHistCnt:= 0;
	xStarted:= FALSE;
	rLatch:= 0.0;
	xLatchValid:= FALSE;
	rSigma:= 0.0;
	xSigmaValid:= FALSE;
	iConsec:= 0;
	iQuar:= 0;
	iHold:= 0;
	iJudgedCnt:= 0;
	iAllDevCnt:= 0;
	xOscOn:= FALSE;
	udiIdxNext:= 0;
	iQdqCnt:= 0;(*分辨率窗一并清空(工况切换)|Yang.zj 2026.10.27+*)
	xPvalValid:= FALSE;
END_IF

(*==================== 丢失帧:不喂模块,原样直通 ====================*)
IF i_xLost THEN
	o_iErrResult:= i_iErr;
	o_byJudge:= 6;(*丢失:没测到不算飞点,锁存不占位*)
	o_xFake:= FALSE;
	RETURN;
END_IF

(*==================== 非新帧周期:全部输出保持上一帧 ====================*)
IF NOT i_xErrValid THEN
	o_iErrResult:= o_iErrResult;
	o_byJudge:= o_byJudge;
	o_xFake:= o_xFake;
	RETURN;
END_IF

byJudge:= 1;(*好,默认*)
rX:= INT_TO_REAL(i_iErr);

udiIdx:= udiIdxNext;
udiIdxNext:= udiIdxNext + 1;

(*==================== 0.数据分辨率quantum:近16个非零相邻差分最小值 ====================*)
(*量化/整数数据上差分MAD可塌缩到0->门限约0,台阶式漂移被判飞点爬行;以分辨率兜底后
 *门限>=5x分辨率,台阶漂移交回趋势带原生跟随;取min对大差分(飞点)免疫,滑窗自适应;
 *连续噪声数据quantum约0不起作用|Yang.zj 2026.10.27+*)
IF xPvalValid AND (udiIdx = udiPidx + 1) THEN(*仅相邻帧的差分入分辨率,跨丢失段不作数*)
	rTmp:= ABS(rX - rPval);
	IF rTmp > 0.0 THEN
		IF iQdqCnt >= 16 THEN
			FOR i:= 0 TO 14 DO
				arQdq[i]:= arQdq[i+1];
			END_FOR
			iQdqCnt:= 15;
		END_IF
		arQdq[iQdqCnt]:= rTmp;
		iQdqCnt:= iQdqCnt + 1;
	END_IF
END_IF
rPval:= rX;
udiPidx:= udiIdx;
xPvalValid:= TRUE;
xQuantumValid:= (iQdqCnt >= 2);
IF xQuantumValid THEN
	rQuantum:= arQdq[0];
	FOR i:= 1 TO iQdqCnt-1 DO
		IF arQdq[i] < rQuantum THEN
			rQuantum:= arQdq[i];
		END_IF
	END_FOR
END_IF

(*==================== 启动期:前2帧无条件采信 ====================*)
IF NOT xStarted THEN
	(*--- 值进可信历史并刷新差分rSigma ---*)
	IF iHistCnt >= KS_FLY_NOISE_WIN THEN
		FOR i:= 0 TO KS_FLY_NOISE_WIN-2 DO
			arHistVal[i]:= arHistVal[i+1];
			auiHistIdx[i]:= auiHistIdx[i+1];
		END_FOR
		iHistCnt:= KS_FLY_NOISE_WIN - 1;
	END_IF
	arHistVal[iHistCnt]:= rX;
	auiHistIdx[iHistCnt]:= udiIdx;
	iHistCnt:= iHistCnt + 1;
	m:= iHistCnt - 1;
	IF m >= KS_FLY_DIFF_MIN THEN
		FOR i:= 0 TO m-1 DO
			arDiff[i]:= arHistVal[i+1] - arHistVal[i];
		END_FOR
		rMed:= KS_FlyMedian(ADR(arDiff), m);
		FOR i:= 0 TO m-1 DO
			arDiff[i]:= ABS(arDiff[i] - rMed);
		END_FOR
		rMed:= KS_FLY_MAD_C / KS_FLY_SQRT2 * KS_FlyMedian(ADR(arDiff), m);
		IF rMed > KS_FLY_EPS THEN
			rSigma:= rMed;
		ELSE
			rSigma:= KS_FLY_EPS;
		END_IF
		xSigmaValid:= TRUE;
	END_IF
	(*--- end push ---*)
	rLatch:= rX;
	xLatchValid:= TRUE;
	IF iHistCnt >= 2 THEN
		xStarted:= TRUE;
	END_IF
	o_iErrResult:= i_iErr;
	o_byJudge:= 0;(*首帧*)
	o_xFake:= FALSE;
	RETURN;
END_IF

(*==================== 1.趋势带参照,量出带外距离rD ====================*)
n:= KS_FLY_TRUST_WIN;
IF iHistCnt < n THEN
	n:= iHistCnt;
END_IF
IF n <= 1 THEN(*阶跃重建后的单点历史:带退化为该点*)
	rA:= arHistVal[iHistCnt-1];
	rB:= rA;
	fP:= rA;(*单点时外推P=该点,与Python _band一致(守卫>=3点时用不到)|Yang.zj 2026.10.27+*)
ELSE
	iBase:= iHistCnt - n;
	m:= 0;
	FOR i:= iBase TO iHistCnt-1 DO
		FOR j:= i+1 TO iHistCnt-1 DO
			udiDt:= auiHistIdx[j] - auiHistIdx[i];(*帧号严格递增,dt>0*)
			IF udiDt > 0 THEN
				arSlope[m]:= (arHistVal[j] - arHistVal[i]) / UDINT_TO_REAL(udiDt);
				m:= m + 1;
			END_IF
		END_FOR
	END_FOR
	IF m > 0 THEN
		fV:= KS_FlyMedian(ADR(arSlope), m);
	ELSE
		fV:= 0.0;
	END_IF
	FOR i:= iBase TO iHistCnt-1 DO
		arExt[i-iBase]:= arHistVal[i] + fV * UDINT_TO_REAL(udiIdx - auiHistIdx[i]);
	END_FOR
	fP:= KS_FlyMedian(ADR(arExt), n);(*外推预测P*)
	FOR i:= iBase TO iHistCnt-1 DO
		arExt[i-iBase]:= arHistVal[i];
	END_FOR
	fL:= KS_FlyMedian(ADR(arExt), n);(*近期水平L*)
	IF fP < fL THEN
		rA:= fP;
		rB:= fL;
	ELSE
		rA:= fL;
		rB:= fP;
	END_IF
END_IF
rD:= 0.0;
IF rX < rA THEN
	rD:= rA - rX;
ELSIF rX > rB THEN
	rD:= rX - rB;
END_IF

(*==================== 2.振荡自愈 ====================*)
rRatio:= 0.0;
IF iJudgedCnt > 0 THEN
	iSum:= 0;
	FOR i:= 0 TO iJudgedCnt-1 DO
		iSum:= iSum + abyJudged[i];
	END_FOR
	rRatio:= INT_TO_REAL(iSum) / INT_TO_REAL(iJudgedCnt);
END_IF
IF iJudgedCnt >= KS_FLY_OSC_WIN THEN
	IF (NOT xOscOn) AND (rRatio > KS_FLY_OSC_IN) THEN
		xOscOn:= TRUE;
	ELSIF xOscOn AND (rRatio < KS_FLY_OSC_OUT) THEN
		xOscOn:= FALSE;
	END_IF
END_IF

(*==================== 3.确定rSigma与两道门槛 ====================*)
IF xSigmaValid THEN
	rS:= rSigma;
	(*σ以数据分辨率兜底(此读取点兜底与Python在push写入时兜底可观测等价:σ仅此处被读)
	 *量化/整数数据门限>=5x分辨率,台阶式漂移交回趋势带原生跟随|Yang.zj 2026.10.27+*)
	IF xQuantumValid AND (rQuantum > rS) THEN
		rS:= rQuantum;
	END_IF
	IF rS < KS_FLY_EPS THEN
		rS:= KS_FLY_EPS;
	END_IF
ELSE
	m:= iHistCnt - 1;
	rTmp:= 0.0;
	IF m > 0 THEN
		FOR i:= 0 TO m-1 DO
			arDiff[i]:= ABS(arHistVal[i+1] - arHistVal[i]);
		END_FOR
		rTmp:= KS_FlyMedian(ADR(arDiff), m);
	END_IF
	(*暖机σ同样以分辨率兜底*)
	IF xQuantumValid AND (rQuantum > rTmp) THEN
		rTmp:= rQuantum;
	END_IF
	IF rTmp < KS_FLY_EPS THEN
		rTmp:= KS_FLY_EPS;
	END_IF
	rS:= KS_FLY_SIG_PROV * rTmp;
END_IF
IF xOscOn AND (iAllDevCnt >= 8) THEN
	FOR i:= 0 TO iAllDevCnt-1 DO
		arDev[i]:= arAllDev[i];
	END_FOR
	rTmp:= KS_FLY_MAD_C * KS_FlyMedian(ADR(arDev), iAllDevCnt);
	IF rTmp > rS THEN
		rS:= rTmp;
	END_IF
END_IF
rTOut:= KS_FLY_K * rS;						(*外门槛*)
rTRet:= KS_FLY_RET_FRAC * KS_FLY_K * rS;	(*回归门槛*)

(*==================== 4.判定状态机(按优先级) ====================*)
IF iQuar > 0 THEN
	(*观察期(刚确认过阶跃):过门进历史但输出/锁存仍是旧电平;未过门撤销观察记1次强超门*)
	IF rD <= rTOut THEN
		iQuar:= iQuar - 1;
		(*--- push ---*)
		IF iHistCnt >= KS_FLY_NOISE_WIN THEN
			FOR i:= 0 TO KS_FLY_NOISE_WIN-2 DO
				arHistVal[i]:= arHistVal[i+1];
				auiHistIdx[i]:= auiHistIdx[i+1];
			END_FOR
			iHistCnt:= KS_FLY_NOISE_WIN - 1;
		END_IF
		arHistVal[iHistCnt]:= rX;
		auiHistIdx[iHistCnt]:= udiIdx;
		iHistCnt:= iHistCnt + 1;
		m:= iHistCnt - 1;
		IF m >= KS_FLY_DIFF_MIN THEN
			FOR i:= 0 TO m-1 DO
				arDiff[i]:= arHistVal[i+1] - arHistVal[i];
			END_FOR
			rMed:= KS_FlyMedian(ADR(arDiff), m);
			FOR i:= 0 TO m-1 DO
				arDiff[i]:= ABS(arDiff[i] - rMed);
			END_FOR
			rMed:= KS_FLY_MAD_C / KS_FLY_SQRT2 * KS_FlyMedian(ADR(arDiff), m);
			IF rMed > KS_FLY_EPS THEN
				rSigma:= rMed;
			ELSE
				rSigma:= KS_FLY_EPS;
			END_IF
			xSigmaValid:= TRUE;
		END_IF
		(*--- end push ---*)
		rOut:= rLatch;
		byJudge:= 2;(*好(观察)*)
	ELSE
		iQuar:= 0;
		iConsec:= 1;
		rOut:= rLatch;(*观察失败一律锁存,不用P*)
		byJudge:= 3;(*飞点*)
	END_IF
ELSIF iConsec > 0 THEN
	(*候选期(已出现强异常):迟滞判回归/续强/暂缓*)
	IF rD <= rTRet THEN
		(*明确回到原趋势:此前强超门判定为飞点,本帧按好点*)
		IF iHistCnt >= KS_FLY_NOISE_WIN THEN
			FOR i:= 0 TO KS_FLY_NOISE_WIN-2 DO
				arHistVal[i]:= arHistVal[i+1];
				auiHistIdx[i]:= auiHistIdx[i+1];
			END_FOR
			iHistCnt:= KS_FLY_NOISE_WIN - 1;
		END_IF
		arHistVal[iHistCnt]:= rX;
		auiHistIdx[iHistCnt]:= udiIdx;
		iHistCnt:= iHistCnt + 1;
		m:= iHistCnt - 1;
		IF m >= KS_FLY_DIFF_MIN THEN
			FOR i:= 0 TO m-1 DO
				arDiff[i]:= arHistVal[i+1] - arHistVal[i];
			END_FOR
			rMed:= KS_FlyMedian(ADR(arDiff), m);
			FOR i:= 0 TO m-1 DO
				arDiff[i]:= ABS(arDiff[i] - rMed);
			END_FOR
			rMed:= KS_FLY_MAD_C / KS_FLY_SQRT2 * KS_FlyMedian(ADR(arDiff), m);
			IF rMed > KS_FLY_EPS THEN
				rSigma:= rMed;
			ELSE
				rSigma:= KS_FLY_EPS;
			END_IF
			xSigmaValid:= TRUE;
		END_IF
		rLatch:= rX;
		xLatchValid:= TRUE;
		iConsec:= 0;
		iHold:= 0;
		rOut:= rX;
	ELSIF rD > rTOut THEN
		iHold:= 0;
		iConsec:= iConsec + 1;
		IF iConsec >= KS_FLY_STEP_CONFIRM THEN
			(*连续强超门满确认帧数->确认阶跃:历史重建为新电平单点,锁存不动,rSigma沿用*)
			arHistVal[0]:= rX;
			auiHistIdx[0]:= udiIdx;
			iHistCnt:= 1;
			iConsec:= 0;
			iQuar:= KS_FLY_QUAR_N;
			rOut:= rLatch;
			byJudge:= 5;(*阶跃*)
		ELSE
			(*替换值:账本>=3点且非振荡模式用趋势外推fP(斜坡上比锁存新鲜)并同步刷锁存,否则退回锁存|Yang.zj 2026.10.27+*)
			IF (iHistCnt >= 3) AND (NOT xOscOn) THEN
				rOut:= fP;
				rLatch:= fP;(*刷锁存:后续阶跃确认/观察帧沿同一条趋势线输出,消除台阶*)
			ELSE
				rOut:= rLatch;
			END_IF
			byJudge:= 3;(*飞点*)
		END_IF
	ELSE
		(*迟滞带内:暂缓不等于判死;连续暂缓满KS_FLY_HOLD_MAX帧按正常值吸收*)
		iHold:= iHold + 1;
		IF iHold >= KS_FLY_HOLD_MAX THEN
			IF iHistCnt >= KS_FLY_NOISE_WIN THEN
				FOR i:= 0 TO KS_FLY_NOISE_WIN-2 DO
					arHistVal[i]:= arHistVal[i+1];
					auiHistIdx[i]:= auiHistIdx[i+1];
				END_FOR
				iHistCnt:= KS_FLY_NOISE_WIN - 1;
			END_IF
			arHistVal[iHistCnt]:= rX;
			auiHistIdx[iHistCnt]:= udiIdx;
			iHistCnt:= iHistCnt + 1;
			m:= iHistCnt - 1;
			IF m >= KS_FLY_DIFF_MIN THEN
				FOR i:= 0 TO m-1 DO
					arDiff[i]:= arHistVal[i+1] - arHistVal[i];
				END_FOR
				rMed:= KS_FlyMedian(ADR(arDiff), m);
				FOR i:= 0 TO m-1 DO
					arDiff[i]:= ABS(arDiff[i] - rMed);
				END_FOR
				rMed:= KS_FLY_MAD_C / KS_FLY_SQRT2 * KS_FlyMedian(ADR(arDiff), m);
				IF rMed > KS_FLY_EPS THEN
					rSigma:= rMed;
				ELSE
					rSigma:= KS_FLY_EPS;
				END_IF
				xSigmaValid:= TRUE;
			END_IF
			rLatch:= rX;
			xLatchValid:= TRUE;
			iConsec:= 0;
			iHold:= 0;
			rOut:= rX;
		ELSE
			(*替换值:账本>=3点且非振荡模式用趋势外推fP并同步刷锁存,否则退回锁存|Yang.zj 2026.10.27+*)
			IF (iHistCnt >= 3) AND (NOT xOscOn) THEN
				rOut:= fP;
				rLatch:= fP;
			ELSE
				rOut:= rLatch;
			END_IF
			byJudge:= 4;(*暂缓*)
		END_IF
	END_IF
ELSIF rD <= rTOut THEN
	(*正常态:带内即好,原值输出*)
	IF iHistCnt >= KS_FLY_NOISE_WIN THEN
		FOR i:= 0 TO KS_FLY_NOISE_WIN-2 DO
			arHistVal[i]:= arHistVal[i+1];
			auiHistIdx[i]:= auiHistIdx[i+1];
		END_FOR
		iHistCnt:= KS_FLY_NOISE_WIN - 1;
	END_IF
	arHistVal[iHistCnt]:= rX;
	auiHistIdx[iHistCnt]:= udiIdx;
	iHistCnt:= iHistCnt + 1;
	m:= iHistCnt - 1;
	IF m >= KS_FLY_DIFF_MIN THEN
		FOR i:= 0 TO m-1 DO
			arDiff[i]:= arHistVal[i+1] - arHistVal[i];
		END_FOR
		rMed:= KS_FlyMedian(ADR(arDiff), m);
		FOR i:= 0 TO m-1 DO
			arDiff[i]:= ABS(arDiff[i] - rMed);
		END_FOR
		rMed:= KS_FLY_MAD_C / KS_FLY_SQRT2 * KS_FlyMedian(ADR(arDiff), m);
		IF rMed > KS_FLY_EPS THEN
			rSigma:= rMed;
		ELSE
			rSigma:= KS_FLY_EPS;
		END_IF
		xSigmaValid:= TRUE;
	END_IF
	rLatch:= rX;
	xLatchValid:= TRUE;
	iConsec:= 0;
	iHold:= 0;
	rOut:= rX;
ELSE
	(*记1次强超门(下一帧来对质)*)
	iConsec:= 1;
	(*替换值:账本>=3点且非振荡模式用趋势外推fP并同步刷锁存,否则退回锁存|Yang.zj 2026.10.27+*)
	IF (iHistCnt >= 3) AND (NOT xOscOn) THEN
		rOut:= fP;
		rLatch:= fP;
	ELSE
		rOut:= rLatch;
	END_IF
	byJudge:= 3;(*飞点*)
END_IF

(*==================== 5.帧末记账(供振荡检测) ====================*)
IF iJudgedCnt >= KS_FLY_OSC_WIN THEN
	FOR i:= 0 TO KS_FLY_OSC_WIN-2 DO
		abyJudged[i]:= abyJudged[i+1];
	END_FOR
	iJudgedCnt:= KS_FLY_OSC_WIN - 1;
END_IF
IF (byJudge <> 1) AND (byJudge <> 2) THEN
	abyJudged[iJudgedCnt]:= 1;
ELSE
	abyJudged[iJudgedCnt]:= 0;
END_IF
iJudgedCnt:= iJudgedCnt + 1;

IF iAllDevCnt >= 16 THEN
	FOR i:= 0 TO 14 DO
		arAllDev[i]:= arAllDev[i+1];
	END_FOR
	iAllDevCnt:= 15;
END_IF
arAllDev[iAllDevCnt]:= ABS(rX - (rA + rB) * 0.5);
iAllDevCnt:= iAllDevCnt + 1;

(*==================== 输出(四舍五入到丝) ====================*)
o_byJudge:= byJudge;
o_xFake:= (byJudge = 3) OR (byJudge = 4);
o_iErrResult:= REAL_TO_INT(rOut);

(* ---- PLC_PRG.st ---- *)
(*@CES
Name=PLC_PRG
Type=FunctionBlock
TypeGuid=6f9dac99-8de1-4efc-8465-68ac443b7d08
Guid=0004b05b-52ec-439c-9f50-4a8655be5d9d
HasDeclaration=True
HasImplementation=True
*)
{DECLARATION}
PROGRAM PLC_PRG
(*主任务-10ms，用于处理弧面信号/套色误差处理等动作*)
VAR
	tiPLC_PRG_Start : TIME;
	tiFunctionEndTime : TIME;
	tiFunctionStartTime : TIME;

	tTime_WriteFileParam_Log: TIME:= T#20S;
	tTime_Cur: TIME;
	tTime_Start_Log: TIME;
	xInitTime_Log: BOOL;

	aiAlarm_V: ARRAY [1..MAX_UNIT_NUM] OF INT;
	aiAlarm_H: ARRAY [1..MAX_UNIT_NUM] OF INT;
	aiAdj_V: ARRAY [1..MAX_UNIT_NUM] OF INT;
	aiAdj_H: ARRAY [1..MAX_UNIT_NUM] OF INT;
	abyAverageNum_V: ARRAY [1..MAX_UNIT_NUM] OF BYTE;
	abyAverageNum_H: ARRAY [1..MAX_UNIT_NUM] OF BYTE;
	//2026.04.11.152628+
	abyAverageNum_Display: ARRAY [1..MAX_UNIT_NUM] OF BYTE;
	astStErrParam_Use: ARRAY [1..MAX_UNIT_NUM] OF StErrParam_Use;
	iN: INT;
	iNum: INT;
	iGrpId: INT;
	xRequstRdAgainOfRingNetDetails: BOOL;

	xInit: BOOL;
	abyLastIndex: ARRAY [1..MAX_UNIT_NUM] OF BYTE;

	(*2025.8.6.193356-套色调整相关*)
	xIsContinue: BOOL;
	axUseErrTransfer: ARRAY [1..2] OF BOOL;
	axCanCalcArcAdjustValue_Grp: ARRAY [1..2] OF BOOL;(*系的计算调整量总标志@控制小黄的耦合算法执行*)
	axCanCalcArcAdjustValue:ARRAY [1..MAX_UNIT_NUM] OF BOOL;
	xRtn: BOOL;
	adwGetArcErrorAxisIdBitIndex: ARRAY [1..2] OF DWORD;(*/.0 轴1 /.1 轴2 ...以此类推*)
	aiGetAxisArcErrorNum: ARRAY [1..2] OF INT;
	dwTempVal: DWORD;
	iStationId: INT;
	iAxisTypeId: INT;
	iUnitId: INT;(*色组号*)

	(*2024.8.1.120147 横向补偿使用的裁切标志*)
	axFlagCutDne_UseHorCompensate_Uw: ARRAY [2..16] OF BOOL;
	axFlagCutDne_UseHorCompensate_Rw: ARRAY [2..16] OF BOOL;
	aiFinalAdjust_V: ARRAY [1..MAX_UNIT_NUM] OF INT;
	aiFinalAdjust_H: ARRAY [1..MAX_UNIT_NUM] OF INT;
	arFinalAdjust_V_ArcList: ARRAY [1..MAX_UNIT_NUM] OF REAL;(*索引为色序的调整量数组*)
	arFinalAdjust_V_Act: ARRAY [1..MAX_UNIT_NUM] OF REAL;(*实际调整量数组*)
	arFinalAdjust_V_Act_ArcList: ARRAY [1..MAX_UNIT_NUM] OF REAL;(*索引为色序的调整量数组*)
	(*2024.7.26.161051 接料补偿@按照每个色组*)
	aiArcActErr_V: ARRAY [2..16] OF INT;(*套色的实际误差@2024.7.26.160439*)
	arD_hat:ARRAY [2..16] OF REAL;(*扰动估计量*)
	(*套色误差使用低通@2024.05.25.132905*)
	arEk_ArcErr_Lp		:ARRAY [2..16,1..3] OF REAL;(*输入寄存器*)
	arE_DEAL_ArcErr_Lp	:ARRAY [2..16,1..3] OF REAL;(*输出寄存器*)
	aiHerror_FollowBefore:ARRAY [1..MAX_UNIT_NUM] OF INT;
	wParam: WORD; (* 丢失|飞点|让料头 *)
	xFlagAdjEnaCalc: BOOL; (* 调整计算使能 *)
	xFlagVelCtl: BOOL; (* 速度控制状态 *)
	lrMaxAdjustVal: LREAL := 0; (* 单周期内最大的调整量 *)
	lrMaxAdjustVal_H: LREAL;		(*2023.6.19.163047*)
	iTmp_DataIndex: INT; (* 误差传递 *)
	iTmp_PrevAxisId: INT; (* 误差传递 *)
	iTmp_RelayErrData_V: INT; (* 误差传递| *)
	iM: INT;
	iSaveTmp_RelayErrData_V: INT;		(*存储的误差传递值*)
	iErForCalc_v: INT; (* 2018.8.22.173310|误差传递| *)
	iError_Curve_Temp_V: INT;
	rError_Curve_Temp_V_Filter: REAL;
	iFinalError_V: INT; (* 纵向最终误差 *)
	iFinalError_H: INT; (* 横向最终误差 *)
	lrTotalAdjustValue: LREAL;		(*总的调整量-实际电机执行的*)
	iFinalAdjust_V: INT; (* 纵向最终调整量 *)
	iFinalAdjust_H: INT; (* 横向最终调整量 *)
	iKp_InUse: INT;
	iKi_InUse: INT;
	iKd_InUse: INT;
	xByPassDeCouple: BOOL;(*跳过解耦控制器*)
	astStArcCoupleRegister:ARRAY [1..2] OF StArcCoupleRegister;(*寄存器参数|索引为系索引*)
	astStArcCoupleRegister_Follow1: ARRAY [1..2] OF StArcCoupleRegister_Follow1;
	byCurGrpId: BYTE;
	arFilmLenth_ArcList: ARRAY [1..DECOUPLD_DDPD_MAX] OF REAL;(*色组的料膜长度@索引为色序-单位mm*)
	rTs: REAL;
	xClrSts: BOOL;
	arDeltaAcceleration_Cur_Delay: ARRAY [2..16,1..20] OF REAL;
	arAcceleration: ARRAY [2..16,1..5] OF REAL;
	arAcceleration_Last:ARRAY [2..16] OF REAL;
	abyAccDecCompensate: ARRAY [2..16] OF BYTE(*=1 补偿开始|=2 补偿结束处理|=0不补偿*);
	arArcVel_LastCycle: ARRAY [2..16,1..2] OF REAL;(*前2拍的速度值|采样周期是圈|[1] 是上一拍,[2]是上上一拍*)
	axDelayCntEn: ARRAY [2..16] OF BOOL;
	abyDelayCnt: ARRAY [2..16] OF BYTE;
	arTarVel_AccDec: ARRAY [2..16] OF REAL;
	arVel_AccelerationEnd: ARRAY [2..16] OF REAL;
	arPrevCycleAcceleration: ARRAY [2..16] OF REAL;(*上一圈的加速度值|用来计算变化量*)
	arPrevCycleDeltaAcceleration: ARRAY [2..16] OF REAL;(*上一拍的加速变化量值@用于判断加速度变化量*)
	axTargetValueTo0_En: ARRAY [2..16] OF BOOL;
	auiCnt_TargetValueTo0_En: ARRAY [2..16] OF UINT;(*使能标志时机计数*)
	arTime_TargetValueTo_ms: ARRAY [2..16] OF REAL;(*目标值到0的时候@ms*)
	arTargetValue_Cur: ARRAY [2..16] OF REAL;
	atPrevCycleTime:ARRAY [2..16] OF TIME;
	arResult_EvenAccSeg:ARRAY [2..16,1..2] OF REAL;

	sFileName_Param: STRING:= FNAME_SYS_PARAM_A;
	iRtn: INT;
	xStartUp: BOOL;

	parCompensateDelayArr: POINTER TO ARRAY [1..200] OF REAL;
	pstStUnitParam_Save: POINTER TO StUnitParam_Save;
	pstStUnitParam_UnSave: POINTER TO StUnitParam_UnSave;
	pstStGrpParam_Save: POINTER TO StGrpParam_Save;
	pstStGrpParam_UnSave: POINTER TO StGrpParam_UnSave;

	//pfbFilter: POINTER TO KS_FB_FiltByAver;(*定义一个只想滤波器的指针*)
	fbKS_FB_GetError_Arc: KS_FB_GetError_Arc;
	afbKS_FB_ARC_PIDAdjust: ARRAY [1..MAX_UNIT_NUM] OF KS_FB_ARC_PIDAdjust;
	fbKS_FB_GetRingNetStationDetails: KS_FB_GetRingNetStationDetails;
	fbKS_FB_StRecord_A: KS_FB_StRecord_A;
//2026.5.9.111535调整量输出放20ms任务吧
//	afbKS_FB_AdjOutCtl: ARRAY [1..2] OF KS_FB_AdjOutCtl;
	iGrp: INT;
	aiGrpAxisList: ARRAY [1..MAX_UNIT_NUM] OF INT; (*系的轴列表*)
	aiStepAdj: ARRAY [1..MAX_UNIT_NUM] OF INT;
	afbKS_FB_VertAdjustCtrl: ARRAY [1..2] OF KS_FB_VertAdjustCtrl;

	uiGroupStationNum: UINT;
	adwInfo_Station: ARRAY [1..128] OF DWORD;
	tmTestSa: TIME;
	tmValue: TIME;

	fbKS_FB_IOConfig: KS_FB_IOConfig;
	fbKS_FB_StepDriveCTL : KS_FB_StepDriveCTL ;
	fbKS_AbsEncModule_IODeal:KS_AbsEncModule_IODeal;
	afbKS_FB_GrpHorzAdjustCtrl:ARRAY [1..2] OF KS_FB_GrpHorzAdjustCtrl;(*横向*)
	iRtn_GetGroupInf: INT;
	aliTime_Value: ARRAY [1..20] OF LTIME;
	iCoreId_1: INT:=1;
	iCoreId_2: INT:=2;
	aiRtn: ARRAY [1..40] OF INT;
	sMsg: STRING;
	iRtn_RdCfg: INT;
	iRtn_WrCfg: INT;

	iMaxRetryTimes: INT := 3;
	aiRetryCount: ARRAY [1..40] OF INT := [0];

	apData : ARRAY [1..MAX_UNIT_NUM] OF UINT;
	apData1 : ARRAY [1..MAX_UNIT_NUM] OF LREAL;
	apData2 : ARRAY [1..MAX_UNIT_NUM] OF LREAL;
	//2025.11.16.104641 跟一色解耦
	afbKS_FB_GetCouplingValue_V:ARRAY [1..2] OF KS_FB_GetCouplingValue_V;
	arCouplingValue: ARRAY [1..MAX_UNIT_NUM] OF REAL;(*索引为色序的调整量数组*)

	aliTime : ARRAY [1..10] OF LTIME;

	aiPress_Manu: ARRAY [1..MAX_UNIT_NUM] OF INT;
	aiUnPress_Manu: ARRAY [1..MAX_UNIT_NUM] OF INT;

	fbKS_FB_GNS_IOCtl: KS_FB_GNS_IOCtl;
	adiGNSIO_Input: ARRAY [1..2] OF DINT;
	diGNSIO_Output: DINT;

	//2026.4.12.134511增加放料弧面检测
	axSensor_Reflex: ARRAY [1..2] OF BOOL;
	iId_Uw_IO: INT;
	iId_Rw_IO: INT;
	iId_If_IO: INT;
	iId_Of_IO: INT;
	axCutCtlEn: ARRAY [1..2] OF BOOL;
	arDiam_NewVol_Use: ARRAY [1..2] OF REAL;
	arVel_Predrv_Use: ARRAY [1..2] OF REAL;
	afbKS_FB_CutDelay_CTL_Uw: ARRAY [1..2] OF KS_FB_CutDelay_CTL_Uw;
	afbTon_DelayTimer_CutOffKnifeCylinder_Uw: ARRAY [1..2] OF TON;
	afbTrig_DelayTimer_CutOffKnifeCylinder_Uw: ARRAY [1..2] OF R_TRIG;//2026.05.25.154820+ 需要一个沿
	axOutput_CutCylinder: ARRAY [1..2] OF BOOL;
	aiCutTotalTime: ARRAY [1..2] OF INT;
	aiDelayMsec_CutOffKnifeCylinder_Final: ARRAY [1..2] OF INT;
	axTorqueCancel: ARRAY [1..2] OF BOOL;
	aiDelayMsec_RollerCylinder_Final: ARRAY [1..2] OF INT;
	aiTimeCnt: ARRAY [1..2] OF INT;
	afbRTrig_Sts_Precuting: ARRAY [1..2] OF R_TRIG;
	axNeedTorqueCancel: ARRAY [1..2] OF BOOL;
	axAxisATorqueCancel_Out: ARRAY [1..2] OF BOOL;
	axAxisBTorqueCancel_Out: ARRAY [1..2] OF BOOL;

//2026.5.8.115201
	hsMode : INT;
	interval : LREAL;
	readHsEnable : INT;

(*月光宝盒异站配置*)
	xRemoteSetDne : BOOL;
	iRemoteSetFailed : INT;
	axRemoteSetDne				: ARRAY [1..MAX_STATION_NUM] OF  BOOL;
	axRemotSetFailed			: ARRAY [1..MAX_STATION_NUM] OF BOOL;

	adwMotorEncoder : ARRAY [1..MAX_UNIT_NUM] OF DWORD := [MAX_UNIT_NUM(4194304)];

	auiAllowMotorRpm_Max : ARRAY [1..MAX_UNIT_NUM] OF UINT := [MAX_UNIT_NUM(5000)];

	udiAddrRd:UDINT;

	iK: INT;
	fbKS_FB_TRIG: R_TRIG;
	xFlag_Stop_Sys: BOOL;//整机系统停机状态
END_VAR

{IMPLEMENTATION}
tiPLC_PRG_Start := TIME();
KS_TskCycle_Begin(ADR(g_astStTaskCycleDetection[1]));

CASE g_iRunStepId OF
	RUNSTEP_STARTUP:
		g_xRunNormalTask:= FALSE;
		Action_StartUp();
		IF xStartUp THEN
			g_iRunStepId:= RUNSTEP_RdRingNetStationDetails;//RUNSTEP_NormalWork;(* 再去加载系统配置文件 *)
		END_IF
	RUNSTEP_RdRingNetStationDetails:
		Action_GetGroupInf();
		g_iRunStepId:= RUNSTEP_LoadSysParam;
	RUNSTEP_LoadSysParam:
		Action_LoadSysParam();
	RUNSTEP_LoadCfg_Motor:
		Action_LoadConfig_Motor();
	RUNSTEP_LoadSysCfg:
		Action_LoadSysCfg();
	RUNSTEP_UpdateSysCfg:
		Action_UpdateSysCfg();
	RUNSTEP_NormalWork:
		g_xRunNormalTask:= TRUE;
		Action_NormalWork();
	RUNSTEP_RESERVED:
		Action_SetSysCfg();
END_CASE

tiFunctionEndTime := TIME();
g_aiFunctionConsueTime[5] := TIME_TO_INT(tiFunctionEndTime-tiFunctionStartTime);

(*主程序逻辑控制结束end-----------------------------*)
(*g_dwPlcLoad:= SysGetPlcLoad(0);(* cpu消耗 *)*)
KS_TskCycle_End(ADR(g_astStTaskCycleDetection[1]));

g_iTime_Main_Task := TIME_TO_INT(TIME()-tiPLC_PRG_Start);

aliTime[10] := aliTime[2] - aliTime[1];
aliTime[9] := aliTime[3] - aliTime[2];
aliTime[8] := aliTime[4] - aliTime[3];
